(* IEC 61131-3 sources: REFUSR/GP/Refusr.jl/samples (part 4) *)

(* ---- 3-MUX_fives-maven-study.st ---- *)
(*
This code implements a shuffled multiplexer with 3 control bits.
The control bits are: Data[6], Data[2], Data[1]
The input bits are: Data[5], Data[7], Data[8], Data[10], Data[11], Data[9], Data[3], Data[4]

The symbolic expression is:
(((((((~((~(D[6]) & ~(D[2])) & ~(D[1])) | D[5]) & (~((D[6] & ~(D[2])) & ~(D[1])) | D[7])) & (~((~(D[6]) & D[2]) & ~(D[1])) | D[8])) & (~((D[6] & D[2]) & ~(D[1])) | D[10])) & (~((~(D[6]) & ~(D[2])) & D[1]) | D[11])) & (~((D[6] & ~(D[2])) & D[1]) | D[9])) & (~((~(D[6]) & D[2]) & D[1]) | D[3])) & (~((D[6] & D[2]) & D[1]) | D[4])

*)

FUNCTION_BLOCK F_CollectInput
  VAR_IN_OUT
      Data : ARRAY[1..15] OF BOOL;
  END_VAR
  VAR_INPUT
      TICK  : BOOL := 0;
      IN1   : BOOL := 0;
      IN2   : BOOL := 0;
      IN3   : BOOL := 0;
      IN4   : BOOL := 0;
      IN5   : BOOL := 0;
      RESET : BOOL := FALSE;
  END_VAR
  VAR_OUTPUT
      Finished : BOOL;
  END_VAR
  VAR
      j    : USINT := 1;
      tock : BOOL  := 0;
  END_VAR
  IF NOT RESET AND tock = NOT TICK THEN
      Data[j]   := IN1;
      Data[j+1] := IN2;
      Data[j+2] := IN3;
      Data[j+3] := IN4;
      Data[j+4] := IN5;
      j := j + 5;
      tock := TICK;
  ELSE
      j := 1;
      tock := 0;
  END_IF;
  Finished := (j > 15);
END_FUNCTION_BLOCK

PROGRAM Boiler
  VAR
    Data  : ARRAY[1..15] OF BOOL;
    Ready : BOOL;
    CollectInput : F_CollectInput;
  END_VAR
  VAR
    TICK     AT %IX1.0 : BOOL;
    IN1      AT %IX0.3 : BOOL;
    IN2      AT %IX0.4 : BOOL;
    IN3      AT %IX0.5 : BOOL;
    IN4      AT %IX0.6 : BOOL;
    IN5      AT %IX0.7 : BOOL;
    OutReady AT %QX0.0 : BOOL := FALSE;
    FeedNext AT %QX0.1 : BOOL := FALSE;
    Out      AT %QX0.2 : BOOL;
  END_VAR
  CollectInput(TICK:=TICK, IN1:=IN1, IN2:=IN2, IN3:=IN3, IN4:=IN4, IN5:=IN5);
  Ready := CollectInput.Finished;
  FeedNext := 1;
  IF Ready THEN
    Out := (((((((((NOT (((NOT D[6]) AND (NOT D[2])) AND (NOT D[1]))) OR D[5]) AND ((NOT ((D[6] AND (NOT D[2])) AND (NOT D[1]))) OR D[7])) AND ((NOT (((NOT D[6]) AND D[2]) AND (NOT D[1]))) OR D[8])) AND ((NOT ((D[6] AND D[2]) AND (NOT D[1]))) OR D[10])) AND ((NOT (((NOT D[6]) AND (NOT D[2])) AND D[1])) OR D[11])) AND ((NOT ((D[6] AND (NOT D[2])) AND D[1])) OR D[9])) AND ((NOT (((NOT D[6]) AND D[2]) AND D[1])) OR D[3])) AND ((NOT ((D[6] AND D[2]) AND D[1])) OR D[4]));
    OutReady := 1;
    CollectInput(RESET:=TRUE);
  END_IF;
END_PROGRAM

CONFIGURATION Config0
  RESOURCE Res0 ON PLC
    TASK task0(INTERVAL := T#20ms,PRIORITY := 0);
    PROGRAM instance0 WITH task0 : Boiler;
  END_RESOURCE
END_CONFIGURATION

(* ---- 3-MUX_flout-chows-peers.st ---- *)
(*
This code implements a shuffled multiplexer with 3 control bits.
The control bits are: Data[1], Data[2], Data[7]
The input bits are: Data[8], Data[3], Data[5], Data[4], Data[9], Data[6], Data[10], Data[11]

The symbolic expression is:
(((((((~((~(D[1]) & ~(D[2])) & ~(D[7])) | D[8]) & (~((D[1] & ~(D[2])) & ~(D[7])) | D[3])) & (~((~(D[1]) & D[2]) & ~(D[7])) | D[5])) & (~((D[1] & D[2]) & ~(D[7])) | D[4])) & (~((~(D[1]) & ~(D[2])) & D[7]) | D[9])) & (~((D[1] & ~(D[2])) & D[7]) | D[6])) & (~((~(D[1]) & D[2]) & D[7]) | D[10])) & (~((D[1] & D[2]) & D[7]) | D[11])

*)

FUNCTION_BLOCK F_CollectInput
  VAR_IN_OUT
      Data : ARRAY[1..15] OF BOOL;
  END_VAR
  VAR_INPUT
      TICK  : BOOL := 0;
      IN1   : BOOL := 0;
      IN2   : BOOL := 0;
      IN3   : BOOL := 0;
      IN4   : BOOL := 0;
      IN5   : BOOL := 0;
      RESET : BOOL := FALSE;
  END_VAR
  VAR_OUTPUT
      Finished : BOOL;
  END_VAR
  VAR
      j    : USINT := 1;
      tock : BOOL  := 0;
  END_VAR
  IF NOT RESET AND tock = NOT TICK THEN
      Data[j]   := IN1;
      Data[j+1] := IN2;
      Data[j+2] := IN3;
      Data[j+3] := IN4;
      Data[j+4] := IN5;
      j := j + 5;
      tock := TICK;
  ELSE
      j := 1;
      tock := 0;
  END_IF;
  Finished := (j > 15);
END_FUNCTION_BLOCK

PROGRAM Boiler
  VAR
    Data  : ARRAY[1..15] OF BOOL;
    Ready : BOOL;
    CollectInput : F_CollectInput;
  END_VAR
  VAR
    TICK     AT %IX1.0 : BOOL;
    IN1      AT %IX0.3 : BOOL;
    IN2      AT %IX0.4 : BOOL;
    IN3      AT %IX0.5 : BOOL;
    IN4      AT %IX0.6 : BOOL;
    IN5      AT %IX0.7 : BOOL;
    OutReady AT %QX0.0 : BOOL := FALSE;
    FeedNext AT %QX0.1 : BOOL := FALSE;
    Out      AT %QX0.2 : BOOL;
  END_VAR
  CollectInput(TICK:=TICK, IN1:=IN1, IN2:=IN2, IN3:=IN3, IN4:=IN4, IN5:=IN5);
  Ready := CollectInput.Finished;
  FeedNext := 1;
  IF Ready THEN
    Out := (((((((((NOT (((NOT D[1]) AND (NOT D[2])) AND (NOT D[7]))) OR D[8]) AND ((NOT ((D[1] AND (NOT D[2])) AND (NOT D[7]))) OR D[3])) AND ((NOT (((NOT D[1]) AND D[2]) AND (NOT D[7]))) OR D[5])) AND ((NOT ((D[1] AND D[2]) AND (NOT D[7]))) OR D[4])) AND ((NOT (((NOT D[1]) AND (NOT D[2])) AND D[7])) OR D[9])) AND ((NOT ((D[1] AND (NOT D[2])) AND D[7])) OR D[6])) AND ((NOT (((NOT D[1]) AND D[2]) AND D[7])) OR D[10])) AND ((NOT ((D[1] AND D[2]) AND D[7])) OR D[11]));
    OutReady := 1;
    CollectInput(RESET:=TRUE);
  END_IF;
END_PROGRAM

CONFIGURATION Config0
  RESOURCE Res0 ON PLC
    TASK task0(INTERVAL := T#20ms,PRIORITY := 0);
    PROGRAM instance0 WITH task0 : Boiler;
  END_RESOURCE
END_CONFIGURATION

(* ---- 3-MUX_fluff-masse-darts.st ---- *)
(*
This code implements a shuffled multiplexer with 3 control bits.
The control bits are: Data[3], Data[2], Data[1]
The input bits are: Data[5], Data[4], Data[6], Data[9], Data[7], Data[11], Data[10], Data[8]

The symbolic expression is:
(((((((~((~(D[3]) & ~(D[2])) & ~(D[1])) | D[5]) & (~((D[3] & ~(D[2])) & ~(D[1])) | D[4])) & (~((~(D[3]) & D[2]) & ~(D[1])) | D[6])) & (~((D[3] & D[2]) & ~(D[1])) | D[9])) & (~((~(D[3]) & ~(D[2])) & D[1]) | D[7])) & (~((D[3] & ~(D[2])) & D[1]) | D[11])) & (~((~(D[3]) & D[2]) & D[1]) | D[10])) & (~((D[3] & D[2]) & D[1]) | D[8])

*)

FUNCTION_BLOCK F_CollectInput
  VAR_IN_OUT
      Data : ARRAY[1..15] OF BOOL;
  END_VAR
  VAR_INPUT
      TICK  : BOOL := 0;
      IN1   : BOOL := 0;
      IN2   : BOOL := 0;
      IN3   : BOOL := 0;
      IN4   : BOOL := 0;
      IN5   : BOOL := 0;
      RESET : BOOL := FALSE;
  END_VAR
  VAR_OUTPUT
      Finished : BOOL;
  END_VAR
  VAR
      j    : USINT := 1;
      tock : BOOL  := 0;
  END_VAR
  IF NOT RESET AND tock = NOT TICK THEN
      Data[j]   := IN1;
      Data[j+1] := IN2;
      Data[j+2] := IN3;
      Data[j+3] := IN4;
      Data[j+4] := IN5;
      j := j + 5;
      tock := TICK;
  ELSE
      j := 1;
      tock := 0;
  END_IF;
  Finished := (j > 15);
END_FUNCTION_BLOCK

PROGRAM Boiler
  VAR
    Data  : ARRAY[1..15] OF BOOL;
    Ready : BOOL;
    CollectInput : F_CollectInput;
  END_VAR
  VAR
    TICK     AT %IX1.0 : BOOL;
    IN1      AT %IX0.3 : BOOL;
    IN2      AT %IX0.4 : BOOL;
    IN3      AT %IX0.5 : BOOL;
    IN4      AT %IX0.6 : BOOL;
    IN5      AT %IX0.7 : BOOL;
    OutReady AT %QX0.0 : BOOL := FALSE;
    FeedNext AT %QX0.1 : BOOL := FALSE;
    Out      AT %QX0.2 : BOOL;
  END_VAR
  CollectInput(TICK:=TICK, IN1:=IN1, IN2:=IN2, IN3:=IN3, IN4:=IN4, IN5:=IN5);
  Ready := CollectInput.Finished;
  FeedNext := 1;
  IF Ready THEN
    Out := (((((((((NOT (((NOT D[3]) AND (NOT D[2])) AND (NOT D[1]))) OR D[5]) AND ((NOT ((D[3] AND (NOT D[2])) AND (NOT D[1]))) OR D[4])) AND ((NOT (((NOT D[3]) AND D[2]) AND (NOT D[1]))) OR D[6])) AND ((NOT ((D[3] AND D[2]) AND (NOT D[1]))) OR D[9])) AND ((NOT (((NOT D[3]) AND (NOT D[2])) AND D[1])) OR D[7])) AND ((NOT ((D[3] AND (NOT D[2])) AND D[1])) OR D[11])) AND ((NOT (((NOT D[3]) AND D[2]) AND D[1])) OR D[10])) AND ((NOT ((D[3] AND D[2]) AND D[1])) OR D[8]));
    OutReady := 1;
    CollectInput(RESET:=TRUE);
  END_IF;
END_PROGRAM

CONFIGURATION Config0
  RESOURCE Res0 ON PLC
    TASK task0(INTERVAL := T#20ms,PRIORITY := 0);
    PROGRAM instance0 WITH task0 : Boiler;
  END_RESOURCE
END_CONFIGURATION

(* ---- 3-MUX_ftped-surfs-skein.st ---- *)
(*
This code implements a shuffled multiplexer with 3 control bits.
The control bits are: Data[3], Data[2], Data[5]
The input bits are: Data[4], Data[7], Data[8], Data[1], Data[10], Data[6], Data[9], Data[11]

The symbolic expression is:
(((((((~((~(D[3]) & ~(D[2])) & ~(D[5])) | D[4]) & (~((D[3] & ~(D[2])) & ~(D[5])) | D[7])) & (~((~(D[3]) & D[2]) & ~(D[5])) | D[8])) & (~((D[3] & D[2]) & ~(D[5])) | D[1])) & (~((~(D[3]) & ~(D[2])) & D[5]) | D[10])) & (~((D[3] & ~(D[2])) & D[5]) | D[6])) & (~((~(D[3]) & D[2]) & D[5]) | D[9])) & (~((D[3] & D[2]) & D[5]) | D[11])

*)

FUNCTION_BLOCK F_CollectInput
  VAR_IN_OUT
      Data : ARRAY[1..15] OF BOOL;
  END_VAR
  VAR_INPUT
      TICK  : BOOL := 0;
      IN1   : BOOL := 0;
      IN2   : BOOL := 0;
      IN3   : BOOL := 0;
      IN4   : BOOL := 0;
      IN5   : BOOL := 0;
      RESET : BOOL := FALSE;
  END_VAR
  VAR_OUTPUT
      Finished : BOOL;
  END_VAR
  VAR
      j    : USINT := 1;
      tock : BOOL  := 0;
  END_VAR
  IF NOT RESET AND tock = NOT TICK THEN
      Data[j]   := IN1;
      Data[j+1] := IN2;
      Data[j+2] := IN3;
      Data[j+3] := IN4;
      Data[j+4] := IN5;
      j := j + 5;
      tock := TICK;
  ELSE
      j := 1;
      tock := 0;
  END_IF;
  Finished := (j > 15);
END_FUNCTION_BLOCK

PROGRAM Boiler
  VAR
    Data  : ARRAY[1..15] OF BOOL;
    Ready : BOOL;
    CollectInput : F_CollectInput;
  END_VAR
  VAR
    TICK     AT %IX1.0 : BOOL;
    IN1      AT %IX0.3 : BOOL;
    IN2      AT %IX0.4 : BOOL;
    IN3      AT %IX0.5 : BOOL;
    IN4      AT %IX0.6 : BOOL;
    IN5      AT %IX0.7 : BOOL;
    OutReady AT %QX0.0 : BOOL := FALSE;
    FeedNext AT %QX0.1 : BOOL := FALSE;
    Out      AT %QX0.2 : BOOL;
  END_VAR
  CollectInput(TICK:=TICK, IN1:=IN1, IN2:=IN2, IN3:=IN3, IN4:=IN4, IN5:=IN5);
  Ready := CollectInput.Finished;
  FeedNext := 1;
  IF Ready THEN
    Out := (((((((((NOT (((NOT D[3]) AND (NOT D[2])) AND (NOT D[5]))) OR D[4]) AND ((NOT ((D[3] AND (NOT D[2])) AND (NOT D[5]))) OR D[7])) AND ((NOT (((NOT D[3]) AND D[2]) AND (NOT D[5]))) OR D[8])) AND ((NOT ((D[3] AND D[2]) AND (NOT D[5]))) OR D[1])) AND ((NOT (((NOT D[3]) AND (NOT D[2])) AND D[5])) OR D[10])) AND ((NOT ((D[3] AND (NOT D[2])) AND D[5])) OR D[6])) AND ((NOT (((NOT D[3]) AND D[2]) AND D[5])) OR D[9])) AND ((NOT ((D[3] AND D[2]) AND D[5])) OR D[11]));
    OutReady := 1;
    CollectInput(RESET:=TRUE);
  END_IF;
END_PROGRAM

CONFIGURATION Config0
  RESOURCE Res0 ON PLC
    TASK task0(INTERVAL := T#20ms,PRIORITY := 0);
    PROGRAM instance0 WITH task0 : Boiler;
  END_RESOURCE
END_CONFIGURATION

(* ---- 3-MUX_fugal-tawny-pants.st ---- *)
(*
This code implements a shuffled multiplexer with 3 control bits.
The control bits are: Data[1], Data[2], Data[3]
The input bits are: Data[5], Data[9], Data[8], Data[4], Data[10], Data[6], Data[7], Data[11]

The symbolic expression is:
(((((((~((~(D[1]) & ~(D[2])) & ~(D[3])) | D[5]) & (~((D[1] & ~(D[2])) & ~(D[3])) | D[9])) & (~((~(D[1]) & D[2]) & ~(D[3])) | D[8])) & (~((D[1] & D[2]) & ~(D[3])) | D[4])) & (~((~(D[1]) & ~(D[2])) & D[3]) | D[10])) & (~((D[1] & ~(D[2])) & D[3]) | D[6])) & (~((~(D[1]) & D[2]) & D[3]) | D[7])) & (~((D[1] & D[2]) & D[3]) | D[11])

*)

FUNCTION_BLOCK F_CollectInput
  VAR_IN_OUT
      Data : ARRAY[1..15] OF BOOL;
  END_VAR
  VAR_INPUT
      TICK  : BOOL := 0;
      IN1   : BOOL := 0;
      IN2   : BOOL := 0;
      IN3   : BOOL := 0;
      IN4   : BOOL := 0;
      IN5   : BOOL := 0;
      RESET : BOOL := FALSE;
  END_VAR
  VAR_OUTPUT
      Finished : BOOL;
  END_VAR
  VAR
      j    : USINT := 1;
      tock : BOOL  := 0;
  END_VAR
  IF NOT RESET AND tock = NOT TICK THEN
      Data[j]   := IN1;
      Data[j+1] := IN2;
      Data[j+2] := IN3;
      Data[j+3] := IN4;
      Data[j+4] := IN5;
      j := j + 5;
      tock := TICK;
  ELSE
      j := 1;
      tock := 0;
  END_IF;
  Finished := (j > 15);
END_FUNCTION_BLOCK

PROGRAM Boiler
  VAR
    Data  : ARRAY[1..15] OF BOOL;
    Ready : BOOL;
    CollectInput : F_CollectInput;
  END_VAR
  VAR
    TICK     AT %IX1.0 : BOOL;
    IN1      AT %IX0.3 : BOOL;
    IN2      AT %IX0.4 : BOOL;
    IN3      AT %IX0.5 : BOOL;
    IN4      AT %IX0.6 : BOOL;
    IN5      AT %IX0.7 : BOOL;
    OutReady AT %QX0.0 : BOOL := FALSE;
    FeedNext AT %QX0.1 : BOOL := FALSE;
    Out      AT %QX0.2 : BOOL;
  END_VAR
  CollectInput(TICK:=TICK, IN1:=IN1, IN2:=IN2, IN3:=IN3, IN4:=IN4, IN5:=IN5);
  Ready := CollectInput.Finished;
  FeedNext := 1;
  IF Ready THEN
    Out := (((((((((NOT (((NOT D[1]) AND (NOT D[2])) AND (NOT D[3]))) OR D[5]) AND ((NOT ((D[1] AND (NOT D[2])) AND (NOT D[3]))) OR D[9])) AND ((NOT (((NOT D[1]) AND D[2]) AND (NOT D[3]))) OR D[8])) AND ((NOT ((D[1] AND D[2]) AND (NOT D[3]))) OR D[4])) AND ((NOT (((NOT D[1]) AND (NOT D[2])) AND D[3])) OR D[10])) AND ((NOT ((D[1] AND (NOT D[2])) AND D[3])) OR D[6])) AND ((NOT (((NOT D[1]) AND D[2]) AND D[3])) OR D[7])) AND ((NOT ((D[1] AND D[2]) AND D[3])) OR D[11]));
    OutReady := 1;
    CollectInput(RESET:=TRUE);
  END_IF;
END_PROGRAM

CONFIGURATION Config0
  RESOURCE Res0 ON PLC
    TASK task0(INTERVAL := T#20ms,PRIORITY := 0);
    PROGRAM instance0 WITH task0 : Boiler;
  END_RESOURCE
END_CONFIGURATION

(* ---- 3-MUX_ghost-throw-niche.st ---- *)
(*
This code implements a shuffled multiplexer with 3 control bits.
The control bits are: Data[2], Data[1], Data[3]
The input bits are: Data[6], Data[5], Data[7], Data[9], Data[10], Data[4], Data[8], Data[11]

The symbolic expression is:
(((((((~((~(D[2]) & ~(D[1])) & ~(D[3])) | D[6]) & (~((D[2] & ~(D[1])) & ~(D[3])) | D[5])) & (~((~(D[2]) & D[1]) & ~(D[3])) | D[7])) & (~((D[2] & D[1]) & ~(D[3])) | D[9])) & (~((~(D[2]) & ~(D[1])) & D[3]) | D[10])) & (~((D[2] & ~(D[1])) & D[3]) | D[4])) & (~((~(D[2]) & D[1]) & D[3]) | D[8])) & (~((D[2] & D[1]) & D[3]) | D[11])

*)

FUNCTION_BLOCK F_CollectInput
  VAR_IN_OUT
      Data : ARRAY[1..15] OF BOOL;
  END_VAR
  VAR_INPUT
      TICK  : BOOL := 0;
      IN1   : BOOL := 0;
      IN2   : BOOL := 0;
      IN3   : BOOL := 0;
      IN4   : BOOL := 0;
      IN5   : BOOL := 0;
      RESET : BOOL := FALSE;
  END_VAR
  VAR_OUTPUT
      Finished : BOOL;
  END_VAR
  VAR
      j    : USINT := 1;
      tock : BOOL  := 0;
  END_VAR
  IF NOT RESET AND tock = NOT TICK THEN
      Data[j]   := IN1;
      Data[j+1] := IN2;
      Data[j+2] := IN3;
      Data[j+3] := IN4;
      Data[j+4] := IN5;
      j := j + 5;
      tock := TICK;
  ELSE
      j := 1;
      tock := 0;
  END_IF;
  Finished := (j > 15);
END_FUNCTION_BLOCK

PROGRAM Boiler
  VAR
    Data  : ARRAY[1..15] OF BOOL;
    Ready : BOOL;
    CollectInput : F_CollectInput;
  END_VAR
  VAR
    TICK     AT %IX1.0 : BOOL;
    IN1      AT %IX0.3 : BOOL;
    IN2      AT %IX0.4 : BOOL;
    IN3      AT %IX0.5 : BOOL;
    IN4      AT %IX0.6 : BOOL;
    IN5      AT %IX0.7 : BOOL;
    OutReady AT %QX0.0 : BOOL := FALSE;
    FeedNext AT %QX0.1 : BOOL := FALSE;
    Out      AT %QX0.2 : BOOL;
  END_VAR
  CollectInput(TICK:=TICK, IN1:=IN1, IN2:=IN2, IN3:=IN3, IN4:=IN4, IN5:=IN5);
  Ready := CollectInput.Finished;
  FeedNext := 1;
  IF Ready THEN
    Out := (((((((((NOT (((NOT D[2]) AND (NOT D[1])) AND (NOT D[3]))) OR D[6]) AND ((NOT ((D[2] AND (NOT D[1])) AND (NOT D[3]))) OR D[5])) AND ((NOT (((NOT D[2]) AND D[1]) AND (NOT D[3]))) OR D[7])) AND ((NOT ((D[2] AND D[1]) AND (NOT D[3]))) OR D[9])) AND ((NOT (((NOT D[2]) AND (NOT D[1])) AND D[3])) OR D[10])) AND ((NOT ((D[2] AND (NOT D[1])) AND D[3])) OR D[4])) AND ((NOT (((NOT D[2]) AND D[1]) AND D[3])) OR D[8])) AND ((NOT ((D[2] AND D[1]) AND D[3])) OR D[11]));
    OutReady := 1;
    CollectInput(RESET:=TRUE);
  END_IF;
END_PROGRAM

CONFIGURATION Config0
  RESOURCE Res0 ON PLC
    TASK task0(INTERVAL := T#20ms,PRIORITY := 0);
    PROGRAM instance0 WITH task0 : Boiler;
  END_RESOURCE
END_CONFIGURATION

(* ---- 3-MUX_giant-blocs-dicta.st ---- *)
(*
This code implements a shuffled multiplexer with 3 control bits.
The control bits are: Data[1], Data[3], Data[9]
The input bits are: Data[4], Data[2], Data[6], Data[8], Data[7], Data[5], Data[11], Data[10]

The symbolic expression is:
(((((((~((~(D[1]) & ~(D[3])) & ~(D[9])) | D[4]) & (~((D[1] & ~(D[3])) & ~(D[9])) | D[2])) & (~((~(D[1]) & D[3]) & ~(D[9])) | D[6])) & (~((D[1] & D[3]) & ~(D[9])) | D[8])) & (~((~(D[1]) & ~(D[3])) & D[9]) | D[7])) & (~((D[1] & ~(D[3])) & D[9]) | D[5])) & (~((~(D[1]) & D[3]) & D[9]) | D[11])) & (~((D[1] & D[3]) & D[9]) | D[10])

*)

FUNCTION_BLOCK F_CollectInput
  VAR_IN_OUT
      Data : ARRAY[1..15] OF BOOL;
  END_VAR
  VAR_INPUT
      TICK  : BOOL := 0;
      IN1   : BOOL := 0;
      IN2   : BOOL := 0;
      IN3   : BOOL := 0;
      IN4   : BOOL := 0;
      IN5   : BOOL := 0;
      RESET : BOOL := FALSE;
  END_VAR
  VAR_OUTPUT
      Finished : BOOL;
  END_VAR
  VAR
      j    : USINT := 1;
      tock : BOOL  := 0;
  END_VAR
  IF NOT RESET AND tock = NOT TICK THEN
      Data[j]   := IN1;
      Data[j+1] := IN2;
      Data[j+2] := IN3;
      Data[j+3] := IN4;
      Data[j+4] := IN5;
      j := j + 5;
      tock := TICK;
  ELSE
      j := 1;
      tock := 0;
  END_IF;
  Finished := (j > 15);
END_FUNCTION_BLOCK

PROGRAM Boiler
  VAR
    Data  : ARRAY[1..15] OF BOOL;
    Ready : BOOL;
    CollectInput : F_CollectInput;
  END_VAR
  VAR
    TICK     AT %IX1.0 : BOOL;
    IN1      AT %IX0.3 : BOOL;
    IN2      AT %IX0.4 : BOOL;
    IN3      AT %IX0.5 : BOOL;
    IN4      AT %IX0.6 : BOOL;
    IN5      AT %IX0.7 : BOOL;
    OutReady AT %QX0.0 : BOOL := FALSE;
    FeedNext AT %QX0.1 : BOOL := FALSE;
    Out      AT %QX0.2 : BOOL;
  END_VAR
  CollectInput(TICK:=TICK, IN1:=IN1, IN2:=IN2, IN3:=IN3, IN4:=IN4, IN5:=IN5);
  Ready := CollectInput.Finished;
  FeedNext := 1;
  IF Ready THEN
    Out := (((((((((NOT (((NOT D[1]) AND (NOT D[3])) AND (NOT D[9]))) OR D[4]) AND ((NOT ((D[1] AND (NOT D[3])) AND (NOT D[9]))) OR D[2])) AND ((NOT (((NOT D[1]) AND D[3]) AND (NOT D[9]))) OR D[6])) AND ((NOT ((D[1] AND D[3]) AND (NOT D[9]))) OR D[8])) AND ((NOT (((NOT D[1]) AND (NOT D[3])) AND D[9])) OR D[7])) AND ((NOT ((D[1] AND (NOT D[3])) AND D[9])) OR D[5])) AND ((NOT (((NOT D[1]) AND D[3]) AND D[9])) OR D[11])) AND ((NOT ((D[1] AND D[3]) AND D[9])) OR D[10]));
    OutReady := 1;
    CollectInput(RESET:=TRUE);
  END_IF;
END_PROGRAM

CONFIGURATION Config0
  RESOURCE Res0 ON PLC
    TASK task0(INTERVAL := T#20ms,PRIORITY := 0);
    PROGRAM instance0 WITH task0 : Boiler;
  END_RESOURCE
END_CONFIGURATION

(* ---- 3-MUX_goofy-uncap-recap.st ---- *)
(*
This code implements a shuffled multiplexer with 3 control bits.
The control bits are: Data[2], Data[1], Data[4]
The input bits are: Data[3], Data[5], Data[7], Data[6], Data[9], Data[10], Data[11], Data[8]

The symbolic expression is:
(((((((~((~(D[2]) & ~(D[1])) & ~(D[4])) | D[3]) & (~((D[2] & ~(D[1])) & ~(D[4])) | D[5])) & (~((~(D[2]) & D[1]) & ~(D[4])) | D[7])) & (~((D[2] & D[1]) & ~(D[4])) | D[6])) & (~((~(D[2]) & ~(D[1])) & D[4]) | D[9])) & (~((D[2] & ~(D[1])) & D[4]) | D[10])) & (~((~(D[2]) & D[1]) & D[4]) | D[11])) & (~((D[2] & D[1]) & D[4]) | D[8])

*)

FUNCTION_BLOCK F_CollectInput
  VAR_IN_OUT
      Data : ARRAY[1..15] OF BOOL;
  END_VAR
  VAR_INPUT
      TICK  : BOOL := 0;
      IN1   : BOOL := 0;
      IN2   : BOOL := 0;
      IN3   : BOOL := 0;
      IN4   : BOOL := 0;
      IN5   : BOOL := 0;
      RESET : BOOL := FALSE;
  END_VAR
  VAR_OUTPUT
      Finished : BOOL;
  END_VAR
  VAR
      j    : USINT := 1;
      tock : BOOL  := 0;
  END_VAR
  IF NOT RESET AND tock = NOT TICK THEN
      Data[j]   := IN1;
      Data[j+1] := IN2;
      Data[j+2] := IN3;
      Data[j+3] := IN4;
      Data[j+4] := IN5;
      j := j + 5;
      tock := TICK;
  ELSE
      j := 1;
      tock := 0;
  END_IF;
  Finished := (j > 15);
END_FUNCTION_BLOCK

PROGRAM Boiler
  VAR
    Data  : ARRAY[1..15] OF BOOL;
    Ready : BOOL;
    CollectInput : F_CollectInput;
  END_VAR
  VAR
    TICK     AT %IX1.0 : BOOL;
    IN1      AT %IX0.3 : BOOL;
    IN2      AT %IX0.4 : BOOL;
    IN3      AT %IX0.5 : BOOL;
    IN4      AT %IX0.6 : BOOL;
    IN5      AT %IX0.7 : BOOL;
    OutReady AT %QX0.0 : BOOL := FALSE;
    FeedNext AT %QX0.1 : BOOL := FALSE;
    Out      AT %QX0.2 : BOOL;
  END_VAR
  CollectInput(TICK:=TICK, IN1:=IN1, IN2:=IN2, IN3:=IN3, IN4:=IN4, IN5:=IN5);
  Ready := CollectInput.Finished;
  FeedNext := 1;
  IF Ready THEN
    Out := (((((((((NOT (((NOT D[2]) AND (NOT D[1])) AND (NOT D[4]))) OR D[3]) AND ((NOT ((D[2] AND (NOT D[1])) AND (NOT D[4]))) OR D[5])) AND ((NOT (((NOT D[2]) AND D[1]) AND (NOT D[4]))) OR D[7])) AND ((NOT ((D[2] AND D[1]) AND (NOT D[4]))) OR D[6])) AND ((NOT (((NOT D[2]) AND (NOT D[1])) AND D[4])) OR D[9])) AND ((NOT ((D[2] AND (NOT D[1])) AND D[4])) OR D[10])) AND ((NOT (((NOT D[2]) AND D[1]) AND D[4])) OR D[11])) AND ((NOT ((D[2] AND D[1]) AND D[4])) OR D[8]));
    OutReady := 1;
    CollectInput(RESET:=TRUE);
  END_IF;
END_PROGRAM

CONFIGURATION Config0
  RESOURCE Res0 ON PLC
    TASK task0(INTERVAL := T#20ms,PRIORITY := 0);
    PROGRAM instance0 WITH task0 : Boiler;
  END_RESOURCE
END_CONFIGURATION

(* ---- 3-MUX_grunt-trite-rapid.st ---- *)
(*
This code implements a shuffled multiplexer with 3 control bits.
The control bits are: Data[2], Data[3], Data[7]
The input bits are: Data[6], Data[4], Data[1], Data[9], Data[5], Data[10], Data[8], Data[11]

The symbolic expression is:
(((((((~((~(D[2]) & ~(D[3])) & ~(D[7])) | D[6]) & (~((D[2] & ~(D[3])) & ~(D[7])) | D[4])) & (~((~(D[2]) & D[3]) & ~(D[7])) | D[1])) & (~((D[2] & D[3]) & ~(D[7])) | D[9])) & (~((~(D[2]) & ~(D[3])) & D[7]) | D[5])) & (~((D[2] & ~(D[3])) & D[7]) | D[10])) & (~((~(D[2]) & D[3]) & D[7]) | D[8])) & (~((D[2] & D[3]) & D[7]) | D[11])

*)

FUNCTION_BLOCK F_CollectInput
  VAR_IN_OUT
      Data : ARRAY[1..15] OF BOOL;
  END_VAR
  VAR_INPUT
      TICK  : BOOL := 0;
      IN1   : BOOL := 0;
      IN2   : BOOL := 0;
      IN3   : BOOL := 0;
      IN4   : BOOL := 0;
      IN5   : BOOL := 0;
      RESET : BOOL := FALSE;
  END_VAR
  VAR_OUTPUT
      Finished : BOOL;
  END_VAR
  VAR
      j    : USINT := 1;
      tock : BOOL  := 0;
  END_VAR
  IF NOT RESET AND tock = NOT TICK THEN
      Data[j]   := IN1;
      Data[j+1] := IN2;
      Data[j+2] := IN3;
      Data[j+3] := IN4;
      Data[j+4] := IN5;
      j := j + 5;
      tock := TICK;
  ELSE
      j := 1;
      tock := 0;
  END_IF;
  Finished := (j > 15);
END_FUNCTION_BLOCK

PROGRAM Boiler
  VAR
    Data  : ARRAY[1..15] OF BOOL;
    Ready : BOOL;
    CollectInput : F_CollectInput;
  END_VAR
  VAR
    TICK     AT %IX1.0 : BOOL;
    IN1      AT %IX0.3 : BOOL;
    IN2      AT %IX0.4 : BOOL;
    IN3      AT %IX0.5 : BOOL;
    IN4      AT %IX0.6 : BOOL;
    IN5      AT %IX0.7 : BOOL;
    OutReady AT %QX0.0 : BOOL := FALSE;
    FeedNext AT %QX0.1 : BOOL := FALSE;
    Out      AT %QX0.2 : BOOL;
  END_VAR
  CollectInput(TICK:=TICK, IN1:=IN1, IN2:=IN2, IN3:=IN3, IN4:=IN4, IN5:=IN5);
  Ready := CollectInput.Finished;
  FeedNext := 1;
  IF Ready THEN
    Out := (((((((((NOT (((NOT D[2]) AND (NOT D[3])) AND (NOT D[7]))) OR D[6]) AND ((NOT ((D[2] AND (NOT D[3])) AND (NOT D[7]))) OR D[4])) AND ((NOT (((NOT D[2]) AND D[3]) AND (NOT D[7]))) OR D[1])) AND ((NOT ((D[2] AND D[3]) AND (NOT D[7]))) OR D[9])) AND ((NOT (((NOT D[2]) AND (NOT D[3])) AND D[7])) OR D[5])) AND ((NOT ((D[2] AND (NOT D[3])) AND D[7])) OR D[10])) AND ((NOT (((NOT D[2]) AND D[3]) AND D[7])) OR D[8])) AND ((NOT ((D[2] AND D[3]) AND D[7])) OR D[11]));
    OutReady := 1;
    CollectInput(RESET:=TRUE);
  END_IF;
END_PROGRAM

CONFIGURATION Config0
  RESOURCE Res0 ON PLC
    TASK task0(INTERVAL := T#20ms,PRIORITY := 0);
    PROGRAM instance0 WITH task0 : Boiler;
  END_RESOURCE
END_CONFIGURATION

(* ---- 3-MUX_gully-crink-seams.st ---- *)
(*
This code implements a shuffled multiplexer with 3 control bits.
The control bits are: Data[1], Data[3], Data[4]
The input bits are: Data[5], Data[2], Data[6], Data[8], Data[9], Data[10], Data[7], Data[11]

The symbolic expression is:
(((((((~((~(D[1]) & ~(D[3])) & ~(D[4])) | D[5]) & (~((D[1] & ~(D[3])) & ~(D[4])) | D[2])) & (~((~(D[1]) & D[3]) & ~(D[4])) | D[6])) & (~((D[1] & D[3]) & ~(D[4])) | D[8])) & (~((~(D[1]) & ~(D[3])) & D[4]) | D[9])) & (~((D[1] & ~(D[3])) & D[4]) | D[10])) & (~((~(D[1]) & D[3]) & D[4]) | D[7])) & (~((D[1] & D[3]) & D[4]) | D[11])

*)

FUNCTION_BLOCK F_CollectInput
  VAR_IN_OUT
      Data : ARRAY[1..15] OF BOOL;
  END_VAR
  VAR_INPUT
      TICK  : BOOL := 0;
      IN1   : BOOL := 0;
      IN2   : BOOL := 0;
      IN3   : BOOL := 0;
      IN4   : BOOL := 0;
      IN5   : BOOL := 0;
      RESET : BOOL := FALSE;
  END_VAR
  VAR_OUTPUT
      Finished : BOOL;
  END_VAR
  VAR
      j    : USINT := 1;
      tock : BOOL  := 0;
  END_VAR
  IF NOT RESET AND tock = NOT TICK THEN
      Data[j]   := IN1;
      Data[j+1] := IN2;
      Data[j+2] := IN3;
      Data[j+3] := IN4;
      Data[j+4] := IN5;
      j := j + 5;
      tock := TICK;
  ELSE
      j := 1;
      tock := 0;
  END_IF;
  Finished := (j > 15);
END_FUNCTION_BLOCK

PROGRAM Boiler
  VAR
    Data  : ARRAY[1..15] OF BOOL;
    Ready : BOOL;
    CollectInput : F_CollectInput;
  END_VAR
  VAR
    TICK     AT %IX1.0 : BOOL;
    IN1      AT %IX0.3 : BOOL;
    IN2      AT %IX0.4 : BOOL;
    IN3      AT %IX0.5 : BOOL;
    IN4      AT %IX0.6 : BOOL;
    IN5      AT %IX0.7 : BOOL;
    OutReady AT %QX0.0 : BOOL := FALSE;
    FeedNext AT %QX0.1 : BOOL := FALSE;
    Out      AT %QX0.2 : BOOL;
  END_VAR
  CollectInput(TICK:=TICK, IN1:=IN1, IN2:=IN2, IN3:=IN3, IN4:=IN4, IN5:=IN5);
  Ready := CollectInput.Finished;
  FeedNext := 1;
  IF Ready THEN
    Out := (((((((((NOT (((NOT D[1]) AND (NOT D[3])) AND (NOT D[4]))) OR D[5]) AND ((NOT ((D[1] AND (NOT D[3])) AND (NOT D[4]))) OR D[2])) AND ((NOT (((NOT D[1]) AND D[3]) AND (NOT D[4]))) OR D[6])) AND ((NOT ((D[1] AND D[3]) AND (NOT D[4]))) OR D[8])) AND ((NOT (((NOT D[1]) AND (NOT D[3])) AND D[4])) OR D[9])) AND ((NOT ((D[1] AND (NOT D[3])) AND D[4])) OR D[10])) AND ((NOT (((NOT D[1]) AND D[3]) AND D[4])) OR D[7])) AND ((NOT ((D[1] AND D[3]) AND D[4])) OR D[11]));
    OutReady := 1;
    CollectInput(RESET:=TRUE);
  END_IF;
END_PROGRAM

CONFIGURATION Config0
  RESOURCE Res0 ON PLC
    TASK task0(INTERVAL := T#20ms,PRIORITY := 0);
    PROGRAM instance0 WITH task0 : Boiler;
  END_RESOURCE
END_CONFIGURATION

(* ---- 3-MUX_hexes-rumps-hanks.st ---- *)
(*
This code implements a shuffled multiplexer with 3 control bits.
The control bits are: Data[2], Data[3], Data[1]
The input bits are: Data[4], Data[5], Data[8], Data[7], Data[6], Data[9], Data[11], Data[10]

The symbolic expression is:
(((((((~((~(D[2]) & ~(D[3])) & ~(D[1])) | D[4]) & (~((D[2] & ~(D[3])) & ~(D[1])) | D[5])) & (~((~(D[2]) & D[3]) & ~(D[1])) | D[8])) & (~((D[2] & D[3]) & ~(D[1])) | D[7])) & (~((~(D[2]) & ~(D[3])) & D[1]) | D[6])) & (~((D[2] & ~(D[3])) & D[1]) | D[9])) & (~((~(D[2]) & D[3]) & D[1]) | D[11])) & (~((D[2] & D[3]) & D[1]) | D[10])

*)

FUNCTION_BLOCK F_CollectInput
  VAR_IN_OUT
      Data : ARRAY[1..15] OF BOOL;
  END_VAR
  VAR_INPUT
      TICK  : BOOL := 0;
      IN1   : BOOL := 0;
      IN2   : BOOL := 0;
      IN3   : BOOL := 0;
      IN4   : BOOL := 0;
      IN5   : BOOL := 0;
      RESET : BOOL := FALSE;
  END_VAR
  VAR_OUTPUT
      Finished : BOOL;
  END_VAR
  VAR
      j    : USINT := 1;
      tock : BOOL  := 0;
  END_VAR
  IF NOT RESET AND tock = NOT TICK THEN
      Data[j]   := IN1;
      Data[j+1] := IN2;
      Data[j+2] := IN3;
      Data[j+3] := IN4;
      Data[j+4] := IN5;
      j := j + 5;
      tock := TICK;
  ELSE
      j := 1;
      tock := 0;
  END_IF;
  Finished := (j > 15);
END_FUNCTION_BLOCK

PROGRAM Boiler
  VAR
    Data  : ARRAY[1..15] OF BOOL;
    Ready : BOOL;
    CollectInput : F_CollectInput;
  END_VAR
  VAR
    TICK     AT %IX1.0 : BOOL;
    IN1      AT %IX0.3 : BOOL;
    IN2      AT %IX0.4 : BOOL;
    IN3      AT %IX0.5 : BOOL;
    IN4      AT %IX0.6 : BOOL;
    IN5      AT %IX0.7 : BOOL;
    OutReady AT %QX0.0 : BOOL := FALSE;
    FeedNext AT %QX0.1 : BOOL := FALSE;
    Out      AT %QX0.2 : BOOL;
  END_VAR
  CollectInput(TICK:=TICK, IN1:=IN1, IN2:=IN2, IN3:=IN3, IN4:=IN4, IN5:=IN5);
  Ready := CollectInput.Finished;
  FeedNext := 1;
  IF Ready THEN
    Out := (((((((((NOT (((NOT D[2]) AND (NOT D[3])) AND (NOT D[1]))) OR D[4]) AND ((NOT ((D[2] AND (NOT D[3])) AND (NOT D[1]))) OR D[5])) AND ((NOT (((NOT D[2]) AND D[3]) AND (NOT D[1]))) OR D[8])) AND ((NOT ((D[2] AND D[3]) AND (NOT D[1]))) OR D[7])) AND ((NOT (((NOT D[2]) AND (NOT D[3])) AND D[1])) OR D[6])) AND ((NOT ((D[2] AND (NOT D[3])) AND D[1])) OR D[9])) AND ((NOT (((NOT D[2]) AND D[3]) AND D[1])) OR D[11])) AND ((NOT ((D[2] AND D[3]) AND D[1])) OR D[10]));
    OutReady := 1;
    CollectInput(RESET:=TRUE);
  END_IF;
END_PROGRAM

CONFIGURATION Config0
  RESOURCE Res0 ON PLC
    TASK task0(INTERVAL := T#20ms,PRIORITY := 0);
    PROGRAM instance0 WITH task0 : Boiler;
  END_RESOURCE
END_CONFIGURATION

(* ---- 3-MUX_hived-field-nuked.st ---- *)
(*
This code implements a shuffled multiplexer with 3 control bits.
The control bits are: Data[4], Data[3], Data[7]
The input bits are: Data[9], Data[10], Data[1], Data[2], Data[5], Data[6], Data[11], Data[8]

The symbolic expression is:
(((((((~((~(D[4]) & ~(D[3])) & ~(D[7])) | D[9]) & (~((D[4] & ~(D[3])) & ~(D[7])) | D[10])) & (~((~(D[4]) & D[3]) & ~(D[7])) | D[1])) & (~((D[4] & D[3]) & ~(D[7])) | D[2])) & (~((~(D[4]) & ~(D[3])) & D[7]) | D[5])) & (~((D[4] & ~(D[3])) & D[7]) | D[6])) & (~((~(D[4]) & D[3]) & D[7]) | D[11])) & (~((D[4] & D[3]) & D[7]) | D[8])

*)

FUNCTION_BLOCK F_CollectInput
  VAR_IN_OUT
      Data : ARRAY[1..15] OF BOOL;
  END_VAR
  VAR_INPUT
      TICK  : BOOL := 0;
      IN1   : BOOL := 0;
      IN2   : BOOL := 0;
      IN3   : BOOL := 0;
      IN4   : BOOL := 0;
      IN5   : BOOL := 0;
      RESET : BOOL := FALSE;
  END_VAR
  VAR_OUTPUT
      Finished : BOOL;
  END_VAR
  VAR
      j    : USINT := 1;
      tock : BOOL  := 0;
  END_VAR
  IF NOT RESET AND tock = NOT TICK THEN
      Data[j]   := IN1;
      Data[j+1] := IN2;
      Data[j+2] := IN3;
      Data[j+3] := IN4;
      Data[j+4] := IN5;
      j := j + 5;
      tock := TICK;
  ELSE
      j := 1;
      tock := 0;
  END_IF;
  Finished := (j > 15);
END_FUNCTION_BLOCK

PROGRAM Boiler
  VAR
    Data  : ARRAY[1..15] OF BOOL;
    Ready : BOOL;
    CollectInput : F_CollectInput;
  END_VAR
  VAR
    TICK     AT %IX1.0 : BOOL;
    IN1      AT %IX0.3 : BOOL;
    IN2      AT %IX0.4 : BOOL;
    IN3      AT %IX0.5 : BOOL;
    IN4      AT %IX0.6 : BOOL;
    IN5      AT %IX0.7 : BOOL;
    OutReady AT %QX0.0 : BOOL := FALSE;
    FeedNext AT %QX0.1 : BOOL := FALSE;
    Out      AT %QX0.2 : BOOL;
  END_VAR
  CollectInput(TICK:=TICK, IN1:=IN1, IN2:=IN2, IN3:=IN3, IN4:=IN4, IN5:=IN5);
  Ready := CollectInput.Finished;
  FeedNext := 1;
  IF Ready THEN
    Out := (((((((((NOT (((NOT D[4]) AND (NOT D[3])) AND (NOT D[7]))) OR D[9]) AND ((NOT ((D[4] AND (NOT D[3])) AND (NOT D[7]))) OR D[10])) AND ((NOT (((NOT D[4]) AND D[3]) AND (NOT D[7]))) OR D[1])) AND ((NOT ((D[4] AND D[3]) AND (NOT D[7]))) OR D[2])) AND ((NOT (((NOT D[4]) AND (NOT D[3])) AND D[7])) OR D[5])) AND ((NOT ((D[4] AND (NOT D[3])) AND D[7])) OR D[6])) AND ((NOT (((NOT D[4]) AND D[3]) AND D[7])) OR D[11])) AND ((NOT ((D[4] AND D[3]) AND D[7])) OR D[8]));
    OutReady := 1;
    CollectInput(RESET:=TRUE);
  END_IF;
END_PROGRAM

CONFIGURATION Config0
  RESOURCE Res0 ON PLC
    TASK task0(INTERVAL := T#20ms,PRIORITY := 0);
    PROGRAM instance0 WITH task0 : Boiler;
  END_RESOURCE
END_CONFIGURATION

(* ---- 3-MUX_jeeps-bazar-carry.st ---- *)
(*
This code implements a shuffled multiplexer with 3 control bits.
The control bits are: Data[2], Data[1], Data[4]
The input bits are: Data[6], Data[5], Data[3], Data[7], Data[9], Data[8], Data[10], Data[11]

The symbolic expression is:
(((((((~((~(D[2]) & ~(D[1])) & ~(D[4])) | D[6]) & (~((D[2] & ~(D[1])) & ~(D[4])) | D[5])) & (~((~(D[2]) & D[1]) & ~(D[4])) | D[3])) & (~((D[2] & D[1]) & ~(D[4])) | D[7])) & (~((~(D[2]) & ~(D[1])) & D[4]) | D[9])) & (~((D[2] & ~(D[1])) & D[4]) | D[8])) & (~((~(D[2]) & D[1]) & D[4]) | D[10])) & (~((D[2] & D[1]) & D[4]) | D[11])

*)

FUNCTION_BLOCK F_CollectInput
  VAR_IN_OUT
      Data : ARRAY[1..15] OF BOOL;
  END_VAR
  VAR_INPUT
      TICK  : BOOL := 0;
      IN1   : BOOL := 0;
      IN2   : BOOL := 0;
      IN3   : BOOL := 0;
      IN4   : BOOL := 0;
      IN5   : BOOL := 0;
      RESET : BOOL := FALSE;
  END_VAR
  VAR_OUTPUT
      Finished : BOOL;
  END_VAR
  VAR
      j    : USINT := 1;
      tock : BOOL  := 0;
  END_VAR
  IF NOT RESET AND tock = NOT TICK THEN
      Data[j]   := IN1;
      Data[j+1] := IN2;
      Data[j+2] := IN3;
      Data[j+3] := IN4;
      Data[j+4] := IN5;
      j := j + 5;
      tock := TICK;
  ELSE
      j := 1;
      tock := 0;
  END_IF;
  Finished := (j > 15);
END_FUNCTION_BLOCK

PROGRAM Boiler
  VAR
    Data  : ARRAY[1..15] OF BOOL;
    Ready : BOOL;
    CollectInput : F_CollectInput;
  END_VAR
  VAR
    TICK     AT %IX1.0 : BOOL;
    IN1      AT %IX0.3 : BOOL;
    IN2      AT %IX0.4 : BOOL;
    IN3      AT %IX0.5 : BOOL;
    IN4      AT %IX0.6 : BOOL;
    IN5      AT %IX0.7 : BOOL;
    OutReady AT %QX0.0 : BOOL := FALSE;
    FeedNext AT %QX0.1 : BOOL := FALSE;
    Out      AT %QX0.2 : BOOL;
  END_VAR
  CollectInput(TICK:=TICK, IN1:=IN1, IN2:=IN2, IN3:=IN3, IN4:=IN4, IN5:=IN5);
  Ready := CollectInput.Finished;
  FeedNext := 1;
  IF Ready THEN
    Out := (((((((((NOT (((NOT D[2]) AND (NOT D[1])) AND (NOT D[4]))) OR D[6]) AND ((NOT ((D[2] AND (NOT D[1])) AND (NOT D[4]))) OR D[5])) AND ((NOT (((NOT D[2]) AND D[1]) AND (NOT D[4]))) OR D[3])) AND ((NOT ((D[2] AND D[1]) AND (NOT D[4]))) OR D[7])) AND ((NOT (((NOT D[2]) AND (NOT D[1])) AND D[4])) OR D[9])) AND ((NOT ((D[2] AND (NOT D[1])) AND D[4])) OR D[8])) AND ((NOT (((NOT D[2]) AND D[1]) AND D[4])) OR D[10])) AND ((NOT ((D[2] AND D[1]) AND D[4])) OR D[11]));
    OutReady := 1;
    CollectInput(RESET:=TRUE);
  END_IF;
END_PROGRAM

CONFIGURATION Config0
  RESOURCE Res0 ON PLC
    TASK task0(INTERVAL := T#20ms,PRIORITY := 0);
    PROGRAM instance0 WITH task0 : Boiler;
  END_RESOURCE
END_CONFIGURATION

(* ---- 3-MUX_jumps-pussy-stirs.st ---- *)
(*
This code implements a shuffled multiplexer with 3 control bits.
The control bits are: Data[2], Data[3], Data[1]
The input bits are: Data[4], Data[5], Data[8], Data[6], Data[7], Data[9], Data[11], Data[10]

The symbolic expression is:
(((((((~((~(D[2]) & ~(D[3])) & ~(D[1])) | D[4]) & (~((D[2] & ~(D[3])) & ~(D[1])) | D[5])) & (~((~(D[2]) & D[3]) & ~(D[1])) | D[8])) & (~((D[2] & D[3]) & ~(D[1])) | D[6])) & (~((~(D[2]) & ~(D[3])) & D[1]) | D[7])) & (~((D[2] & ~(D[3])) & D[1]) | D[9])) & (~((~(D[2]) & D[3]) & D[1]) | D[11])) & (~((D[2] & D[3]) & D[1]) | D[10])

*)

FUNCTION_BLOCK F_CollectInput
  VAR_IN_OUT
      Data : ARRAY[1..15] OF BOOL;
  END_VAR
  VAR_INPUT
      TICK  : BOOL := 0;
      IN1   : BOOL := 0;
      IN2   : BOOL := 0;
      IN3   : BOOL := 0;
      IN4   : BOOL := 0;
      IN5   : BOOL := 0;
      RESET : BOOL := FALSE;
  END_VAR
  VAR_OUTPUT
      Finished : BOOL;
  END_VAR
  VAR
      j    : USINT := 1;
      tock : BOOL  := 0;
  END_VAR
  IF NOT RESET AND tock = NOT TICK THEN
      Data[j]   := IN1;
      Data[j+1] := IN2;
      Data[j+2] := IN3;
      Data[j+3] := IN4;
      Data[j+4] := IN5;
      j := j + 5;
      tock := TICK;
  ELSE
      j := 1;
      tock := 0;
  END_IF;
  Finished := (j > 15);
END_FUNCTION_BLOCK

PROGRAM Boiler
  VAR
    Data  : ARRAY[1..15] OF BOOL;
    Ready : BOOL;
    CollectInput : F_CollectInput;
  END_VAR
  VAR
    TICK     AT %IX1.0 : BOOL;
    IN1      AT %IX0.3 : BOOL;
    IN2      AT %IX0.4 : BOOL;
    IN3      AT %IX0.5 : BOOL;
    IN4      AT %IX0.6 : BOOL;
    IN5      AT %IX0.7 : BOOL;
    OutReady AT %QX0.0 : BOOL := FALSE;
    FeedNext AT %QX0.1 : BOOL := FALSE;
    Out      AT %QX0.2 : BOOL;
  END_VAR
  CollectInput(TICK:=TICK, IN1:=IN1, IN2:=IN2, IN3:=IN3, IN4:=IN4, IN5:=IN5);
  Ready := CollectInput.Finished;
  FeedNext := 1;
  IF Ready THEN
    Out := (((((((((NOT (((NOT D[2]) AND (NOT D[3])) AND (NOT D[1]))) OR D[4]) AND ((NOT ((D[2] AND (NOT D[3])) AND (NOT D[1]))) OR D[5])) AND ((NOT (((NOT D[2]) AND D[3]) AND (NOT D[1]))) OR D[8])) AND ((NOT ((D[2] AND D[3]) AND (NOT D[1]))) OR D[6])) AND ((NOT (((NOT D[2]) AND (NOT D[3])) AND D[1])) OR D[7])) AND ((NOT ((D[2] AND (NOT D[3])) AND D[1])) OR D[9])) AND ((NOT (((NOT D[2]) AND D[3]) AND D[1])) OR D[11])) AND ((NOT ((D[2] AND D[3]) AND D[1])) OR D[10]));
    OutReady := 1;
    CollectInput(RESET:=TRUE);
  END_IF;
END_PROGRAM

CONFIGURATION Config0
  RESOURCE Res0 ON PLC
    TASK task0(INTERVAL := T#20ms,PRIORITY := 0);
    PROGRAM instance0 WITH task0 : Boiler;
  END_RESOURCE
END_CONFIGURATION

(* ---- 3-MUX_laves-tidal-green.st ---- *)
(*
This code implements a shuffled multiplexer with 3 control bits.
The control bits are: Data[2], Data[3], Data[1]
The input bits are: Data[5], Data[8], Data[6], Data[4], Data[7], Data[9], Data[10], Data[11]

The symbolic expression is:
(((((((~((~(D[2]) & ~(D[3])) & ~(D[1])) | D[5]) & (~((D[2] & ~(D[3])) & ~(D[1])) | D[8])) & (~((~(D[2]) & D[3]) & ~(D[1])) | D[6])) & (~((D[2] & D[3]) & ~(D[1])) | D[4])) & (~((~(D[2]) & ~(D[3])) & D[1]) | D[7])) & (~((D[2] & ~(D[3])) & D[1]) | D[9])) & (~((~(D[2]) & D[3]) & D[1]) | D[10])) & (~((D[2] & D[3]) & D[1]) | D[11])

*)

FUNCTION_BLOCK F_CollectInput
  VAR_IN_OUT
      Data : ARRAY[1..15] OF BOOL;
  END_VAR
  VAR_INPUT
      TICK  : BOOL := 0;
      IN1   : BOOL := 0;
      IN2   : BOOL := 0;
      IN3   : BOOL := 0;
      IN4   : BOOL := 0;
      IN5   : BOOL := 0;
      RESET : BOOL := FALSE;
  END_VAR
  VAR_OUTPUT
      Finished : BOOL;
  END_VAR
  VAR
      j    : USINT := 1;
      tock : BOOL  := 0;
  END_VAR
  IF NOT RESET AND tock = NOT TICK THEN
      Data[j]   := IN1;
      Data[j+1] := IN2;
      Data[j+2] := IN3;
      Data[j+3] := IN4;
      Data[j+4] := IN5;
      j := j + 5;
      tock := TICK;
  ELSE
      j := 1;
      tock := 0;
  END_IF;
  Finished := (j > 15);
END_FUNCTION_BLOCK

PROGRAM Boiler
  VAR
    Data  : ARRAY[1..15] OF BOOL;
    Ready : BOOL;
    CollectInput : F_CollectInput;
  END_VAR
  VAR
    TICK     AT %IX1.0 : BOOL;
    IN1      AT %IX0.3 : BOOL;
    IN2      AT %IX0.4 : BOOL;
    IN3      AT %IX0.5 : BOOL;
    IN4      AT %IX0.6 : BOOL;
    IN5      AT %IX0.7 : BOOL;
    OutReady AT %QX0.0 : BOOL := FALSE;
    FeedNext AT %QX0.1 : BOOL := FALSE;
    Out      AT %QX0.2 : BOOL;
  END_VAR
  CollectInput(TICK:=TICK, IN1:=IN1, IN2:=IN2, IN3:=IN3, IN4:=IN4, IN5:=IN5);
  Ready := CollectInput.Finished;
  FeedNext := 1;
  IF Ready THEN
    Out := (((((((((NOT (((NOT D[2]) AND (NOT D[3])) AND (NOT D[1]))) OR D[5]) AND ((NOT ((D[2] AND (NOT D[3])) AND (NOT D[1]))) OR D[8])) AND ((NOT (((NOT D[2]) AND D[3]) AND (NOT D[1]))) OR D[6])) AND ((NOT ((D[2] AND D[3]) AND (NOT D[1]))) OR D[4])) AND ((NOT (((NOT D[2]) AND (NOT D[3])) AND D[1])) OR D[7])) AND ((NOT ((D[2] AND (NOT D[3])) AND D[1])) OR D[9])) AND ((NOT (((NOT D[2]) AND D[3]) AND D[1])) OR D[10])) AND ((NOT ((D[2] AND D[3]) AND D[1])) OR D[11]));
    OutReady := 1;
    CollectInput(RESET:=TRUE);
  END_IF;
END_PROGRAM

CONFIGURATION Config0
  RESOURCE Res0 ON PLC
    TASK task0(INTERVAL := T#20ms,PRIORITY := 0);
    PROGRAM instance0 WITH task0 : Boiler;
  END_RESOURCE
END_CONFIGURATION

(* ---- 3-MUX_leers-curse-altho.st ---- *)
(*
This code implements a shuffled multiplexer with 3 control bits.
The control bits are: Data[3], Data[1], Data[2]
The input bits are: Data[4], Data[6], Data[5], Data[7], Data[9], Data[8], Data[11], Data[10]

The symbolic expression is:
(((((((~((~(D[3]) & ~(D[1])) & ~(D[2])) | D[4]) & (~((D[3] & ~(D[1])) & ~(D[2])) | D[6])) & (~((~(D[3]) & D[1]) & ~(D[2])) | D[5])) & (~((D[3] & D[1]) & ~(D[2])) | D[7])) & (~((~(D[3]) & ~(D[1])) & D[2]) | D[9])) & (~((D[3] & ~(D[1])) & D[2]) | D[8])) & (~((~(D[3]) & D[1]) & D[2]) | D[11])) & (~((D[3] & D[1]) & D[2]) | D[10])

*)

FUNCTION_BLOCK F_CollectInput
  VAR_IN_OUT
      Data : ARRAY[1..15] OF BOOL;
  END_VAR
  VAR_INPUT
      TICK  : BOOL := 0;
      IN1   : BOOL := 0;
      IN2   : BOOL := 0;
      IN3   : BOOL := 0;
      IN4   : BOOL := 0;
      IN5   : BOOL := 0;
      RESET : BOOL := FALSE;
  END_VAR
  VAR_OUTPUT
      Finished : BOOL;
  END_VAR
  VAR
      j    : USINT := 1;
      tock : BOOL  := 0;
  END_VAR
  IF NOT RESET AND tock = NOT TICK THEN
      Data[j]   := IN1;
      Data[j+1] := IN2;
      Data[j+2] := IN3;
      Data[j+3] := IN4;
      Data[j+4] := IN5;
      j := j + 5;
      tock := TICK;
  ELSE
      j := 1;
      tock := 0;
  END_IF;
  Finished := (j > 15);
END_FUNCTION_BLOCK

PROGRAM Boiler
  VAR
    Data  : ARRAY[1..15] OF BOOL;
    Ready : BOOL;
    CollectInput : F_CollectInput;
  END_VAR
  VAR
    TICK     AT %IX1.0 : BOOL;
    IN1      AT %IX0.3 : BOOL;
    IN2      AT %IX0.4 : BOOL;
    IN3      AT %IX0.5 : BOOL;
    IN4      AT %IX0.6 : BOOL;
    IN5      AT %IX0.7 : BOOL;
    OutReady AT %QX0.0 : BOOL := FALSE;
    FeedNext AT %QX0.1 : BOOL := FALSE;
    Out      AT %QX0.2 : BOOL;
  END_VAR
  CollectInput(TICK:=TICK, IN1:=IN1, IN2:=IN2, IN3:=IN3, IN4:=IN4, IN5:=IN5);
  Ready := CollectInput.Finished;
  FeedNext := 1;
  IF Ready THEN
    Out := (((((((((NOT (((NOT D[3]) AND (NOT D[1])) AND (NOT D[2]))) OR D[4]) AND ((NOT ((D[3] AND (NOT D[1])) AND (NOT D[2]))) OR D[6])) AND ((NOT (((NOT D[3]) AND D[1]) AND (NOT D[2]))) OR D[5])) AND ((NOT ((D[3] AND D[1]) AND (NOT D[2]))) OR D[7])) AND ((NOT (((NOT D[3]) AND (NOT D[1])) AND D[2])) OR D[9])) AND ((NOT ((D[3] AND (NOT D[1])) AND D[2])) OR D[8])) AND ((NOT (((NOT D[3]) AND D[1]) AND D[2])) OR D[11])) AND ((NOT ((D[3] AND D[1]) AND D[2])) OR D[10]));
    OutReady := 1;
    CollectInput(RESET:=TRUE);
  END_IF;
END_PROGRAM

CONFIGURATION Config0
  RESOURCE Res0 ON PLC
    TASK task0(INTERVAL := T#20ms,PRIORITY := 0);
    PROGRAM instance0 WITH task0 : Boiler;
  END_RESOURCE
END_CONFIGURATION

(* ---- 3-MUX_legos-taker-gauze.st ---- *)
(*
This code implements a shuffled multiplexer with 3 control bits.
The control bits are: Data[2], Data[1], Data[3]
The input bits are: Data[6], Data[5], Data[7], Data[4], Data[8], Data[9], Data[11], Data[10]

The symbolic expression is:
(((((((~((~(D[2]) & ~(D[1])) & ~(D[3])) | D[6]) & (~((D[2] & ~(D[1])) & ~(D[3])) | D[5])) & (~((~(D[2]) & D[1]) & ~(D[3])) | D[7])) & (~((D[2] & D[1]) & ~(D[3])) | D[4])) & (~((~(D[2]) & ~(D[1])) & D[3]) | D[8])) & (~((D[2] & ~(D[1])) & D[3]) | D[9])) & (~((~(D[2]) & D[1]) & D[3]) | D[11])) & (~((D[2] & D[1]) & D[3]) | D[10])

*)

FUNCTION_BLOCK F_CollectInput
  VAR_IN_OUT
      Data : ARRAY[1..15] OF BOOL;
  END_VAR
  VAR_INPUT
      TICK  : BOOL := 0;
      IN1   : BOOL := 0;
      IN2   : BOOL := 0;
      IN3   : BOOL := 0;
      IN4   : BOOL := 0;
      IN5   : BOOL := 0;
      RESET : BOOL := FALSE;
  END_VAR
  VAR_OUTPUT
      Finished : BOOL;
  END_VAR
  VAR
      j    : USINT := 1;
      tock : BOOL  := 0;
  END_VAR
  IF NOT RESET AND tock = NOT TICK THEN
      Data[j]   := IN1;
      Data[j+1] := IN2;
      Data[j+2] := IN3;
      Data[j+3] := IN4;
      Data[j+4] := IN5;
      j := j + 5;
      tock := TICK;
  ELSE
      j := 1;
      tock := 0;
  END_IF;
  Finished := (j > 15);
END_FUNCTION_BLOCK

PROGRAM Boiler
  VAR
    Data  : ARRAY[1..15] OF BOOL;
    Ready : BOOL;
    CollectInput : F_CollectInput;
  END_VAR
  VAR
    TICK     AT %IX1.0 : BOOL;
    IN1      AT %IX0.3 : BOOL;
    IN2      AT %IX0.4 : BOOL;
    IN3      AT %IX0.5 : BOOL;
    IN4      AT %IX0.6 : BOOL;
    IN5      AT %IX0.7 : BOOL;
    OutReady AT %QX0.0 : BOOL := FALSE;
    FeedNext AT %QX0.1 : BOOL := FALSE;
    Out      AT %QX0.2 : BOOL;
  END_VAR
  CollectInput(TICK:=TICK, IN1:=IN1, IN2:=IN2, IN3:=IN3, IN4:=IN4, IN5:=IN5);
  Ready := CollectInput.Finished;
  FeedNext := 1;
  IF Ready THEN
    Out := (((((((((NOT (((NOT D[2]) AND (NOT D[1])) AND (NOT D[3]))) OR D[6]) AND ((NOT ((D[2] AND (NOT D[1])) AND (NOT D[3]))) OR D[5])) AND ((NOT (((NOT D[2]) AND D[1]) AND (NOT D[3]))) OR D[7])) AND ((NOT ((D[2] AND D[1]) AND (NOT D[3]))) OR D[4])) AND ((NOT (((NOT D[2]) AND (NOT D[1])) AND D[3])) OR D[8])) AND ((NOT ((D[2] AND (NOT D[1])) AND D[3])) OR D[9])) AND ((NOT (((NOT D[2]) AND D[1]) AND D[3])) OR D[11])) AND ((NOT ((D[2] AND D[1]) AND D[3])) OR D[10]));
    OutReady := 1;
    CollectInput(RESET:=TRUE);
  END_IF;
END_PROGRAM

CONFIGURATION Config0
  RESOURCE Res0 ON PLC
    TASK task0(INTERVAL := T#20ms,PRIORITY := 0);
    PROGRAM instance0 WITH task0 : Boiler;
  END_RESOURCE
END_CONFIGURATION

(* ---- 3-MUX_loony-spume-duvet.st ---- *)
(*
This code implements a shuffled multiplexer with 3 control bits.
The control bits are: Data[1], Data[2], Data[3]
The input bits are: Data[5], Data[6], Data[10], Data[4], Data[11], Data[7], Data[8], Data[9]

The symbolic expression is:
(((((((~((~(D[1]) & ~(D[2])) & ~(D[3])) | D[5]) & (~((D[1] & ~(D[2])) & ~(D[3])) | D[6])) & (~((~(D[1]) & D[2]) & ~(D[3])) | D[10])) & (~((D[1] & D[2]) & ~(D[3])) | D[4])) & (~((~(D[1]) & ~(D[2])) & D[3]) | D[11])) & (~((D[1] & ~(D[2])) & D[3]) | D[7])) & (~((~(D[1]) & D[2]) & D[3]) | D[8])) & (~((D[1] & D[2]) & D[3]) | D[9])

*)

FUNCTION_BLOCK F_CollectInput
  VAR_IN_OUT
      Data : ARRAY[1..15] OF BOOL;
  END_VAR
  VAR_INPUT
      TICK  : BOOL := 0;
      IN1   : BOOL := 0;
      IN2   : BOOL := 0;
      IN3   : BOOL := 0;
      IN4   : BOOL := 0;
      IN5   : BOOL := 0;
      RESET : BOOL := FALSE;
  END_VAR
  VAR_OUTPUT
      Finished : BOOL;
  END_VAR
  VAR
      j    : USINT := 1;
      tock : BOOL  := 0;
  END_VAR
  IF NOT RESET AND tock = NOT TICK THEN
      Data[j]   := IN1;
      Data[j+1] := IN2;
      Data[j+2] := IN3;
      Data[j+3] := IN4;
      Data[j+4] := IN5;
      j := j + 5;
      tock := TICK;
  ELSE
      j := 1;
      tock := 0;
  END_IF;
  Finished := (j > 15);
END_FUNCTION_BLOCK

PROGRAM Boiler
  VAR
    Data  : ARRAY[1..15] OF BOOL;
    Ready : BOOL;
    CollectInput : F_CollectInput;
  END_VAR
  VAR
    TICK     AT %IX1.0 : BOOL;
    IN1      AT %IX0.3 : BOOL;
    IN2      AT %IX0.4 : BOOL;
    IN3      AT %IX0.5 : BOOL;
    IN4      AT %IX0.6 : BOOL;
    IN5      AT %IX0.7 : BOOL;
    OutReady AT %QX0.0 : BOOL := FALSE;
    FeedNext AT %QX0.1 : BOOL := FALSE;
    Out      AT %QX0.2 : BOOL;
  END_VAR
  CollectInput(TICK:=TICK, IN1:=IN1, IN2:=IN2, IN3:=IN3, IN4:=IN4, IN5:=IN5);
  Ready := CollectInput.Finished;
  FeedNext := 1;
  IF Ready THEN
    Out := (((((((((NOT (((NOT D[1]) AND (NOT D[2])) AND (NOT D[3]))) OR D[5]) AND ((NOT ((D[1] AND (NOT D[2])) AND (NOT D[3]))) OR D[6])) AND ((NOT (((NOT D[1]) AND D[2]) AND (NOT D[3]))) OR D[10])) AND ((NOT ((D[1] AND D[2]) AND (NOT D[3]))) OR D[4])) AND ((NOT (((NOT D[1]) AND (NOT D[2])) AND D[3])) OR D[11])) AND ((NOT ((D[1] AND (NOT D[2])) AND D[3])) OR D[7])) AND ((NOT (((NOT D[1]) AND D[2]) AND D[3])) OR D[8])) AND ((NOT ((D[1] AND D[2]) AND D[3])) OR D[9]));
    OutReady := 1;
    CollectInput(RESET:=TRUE);
  END_IF;
END_PROGRAM

CONFIGURATION Config0
  RESOURCE Res0 ON PLC
    TASK task0(INTERVAL := T#20ms,PRIORITY := 0);
    PROGRAM instance0 WITH task0 : Boiler;
  END_RESOURCE
END_CONFIGURATION

(* ---- 3-MUX_magus-taxol-cones.st ---- *)
(*
This code implements a shuffled multiplexer with 3 control bits.
The control bits are: Data[3], Data[2], Data[4]
The input bits are: Data[1], Data[6], Data[5], Data[8], Data[7], Data[9], Data[10], Data[11]

The symbolic expression is:
(((((((~((~(D[3]) & ~(D[2])) & ~(D[4])) | D[1]) & (~((D[3] & ~(D[2])) & ~(D[4])) | D[6])) & (~((~(D[3]) & D[2]) & ~(D[4])) | D[5])) & (~((D[3] & D[2]) & ~(D[4])) | D[8])) & (~((~(D[3]) & ~(D[2])) & D[4]) | D[7])) & (~((D[3] & ~(D[2])) & D[4]) | D[9])) & (~((~(D[3]) & D[2]) & D[4]) | D[10])) & (~((D[3] & D[2]) & D[4]) | D[11])

*)

FUNCTION_BLOCK F_CollectInput
  VAR_IN_OUT
      Data : ARRAY[1..15] OF BOOL;
  END_VAR
  VAR_INPUT
      TICK  : BOOL := 0;
      IN1   : BOOL := 0;
      IN2   : BOOL := 0;
      IN3   : BOOL := 0;
      IN4   : BOOL := 0;
      IN5   : BOOL := 0;
      RESET : BOOL := FALSE;
  END_VAR
  VAR_OUTPUT
      Finished : BOOL;
  END_VAR
  VAR
      j    : USINT := 1;
      tock : BOOL  := 0;
  END_VAR
  IF NOT RESET AND tock = NOT TICK THEN
      Data[j]   := IN1;
      Data[j+1] := IN2;
      Data[j+2] := IN3;
      Data[j+3] := IN4;
      Data[j+4] := IN5;
      j := j + 5;
      tock := TICK;
  ELSE
      j := 1;
      tock := 0;
  END_IF;
  Finished := (j > 15);
END_FUNCTION_BLOCK

PROGRAM Boiler
  VAR
    Data  : ARRAY[1..15] OF BOOL;
    Ready : BOOL;
    CollectInput : F_CollectInput;
  END_VAR
  VAR
    TICK     AT %IX1.0 : BOOL;
    IN1      AT %IX0.3 : BOOL;
    IN2      AT %IX0.4 : BOOL;
    IN3      AT %IX0.5 : BOOL;
    IN4      AT %IX0.6 : BOOL;
    IN5      AT %IX0.7 : BOOL;
    OutReady AT %QX0.0 : BOOL := FALSE;
    FeedNext AT %QX0.1 : BOOL := FALSE;
    Out      AT %QX0.2 : BOOL;
  END_VAR
  CollectInput(TICK:=TICK, IN1:=IN1, IN2:=IN2, IN3:=IN3, IN4:=IN4, IN5:=IN5);
  Ready := CollectInput.Finished;
  FeedNext := 1;
  IF Ready THEN
    Out := (((((((((NOT (((NOT D[3]) AND (NOT D[2])) AND (NOT D[4]))) OR D[1]) AND ((NOT ((D[3] AND (NOT D[2])) AND (NOT D[4]))) OR D[6])) AND ((NOT (((NOT D[3]) AND D[2]) AND (NOT D[4]))) OR D[5])) AND ((NOT ((D[3] AND D[2]) AND (NOT D[4]))) OR D[8])) AND ((NOT (((NOT D[3]) AND (NOT D[2])) AND D[4])) OR D[7])) AND ((NOT ((D[3] AND (NOT D[2])) AND D[4])) OR D[9])) AND ((NOT (((NOT D[3]) AND D[2]) AND D[4])) OR D[10])) AND ((NOT ((D[3] AND D[2]) AND D[4])) OR D[11]));
    OutReady := 1;
    CollectInput(RESET:=TRUE);
  END_IF;
END_PROGRAM

CONFIGURATION Config0
  RESOURCE Res0 ON PLC
    TASK task0(INTERVAL := T#20ms,PRIORITY := 0);
    PROGRAM instance0 WITH task0 : Boiler;
  END_RESOURCE
END_CONFIGURATION

(* ---- 3-MUX_mazes-villi-eared.st ---- *)
(*
This code implements a shuffled multiplexer with 3 control bits.
The control bits are: Data[8], Data[3], Data[4]
The input bits are: Data[2], Data[1], Data[5], Data[6], Data[7], Data[9], Data[10], Data[11]

The symbolic expression is:
(((((((~((~(D[8]) & ~(D[3])) & ~(D[4])) | D[2]) & (~((D[8] & ~(D[3])) & ~(D[4])) | D[1])) & (~((~(D[8]) & D[3]) & ~(D[4])) | D[5])) & (~((D[8] & D[3]) & ~(D[4])) | D[6])) & (~((~(D[8]) & ~(D[3])) & D[4]) | D[7])) & (~((D[8] & ~(D[3])) & D[4]) | D[9])) & (~((~(D[8]) & D[3]) & D[4]) | D[10])) & (~((D[8] & D[3]) & D[4]) | D[11])

*)

FUNCTION_BLOCK F_CollectInput
  VAR_IN_OUT
      Data : ARRAY[1..15] OF BOOL;
  END_VAR
  VAR_INPUT
      TICK  : BOOL := 0;
      IN1   : BOOL := 0;
      IN2   : BOOL := 0;
      IN3   : BOOL := 0;
      IN4   : BOOL := 0;
      IN5   : BOOL := 0;
      RESET : BOOL := FALSE;
  END_VAR
  VAR_OUTPUT
      Finished : BOOL;
  END_VAR
  VAR
      j    : USINT := 1;
      tock : BOOL  := 0;
  END_VAR
  IF NOT RESET AND tock = NOT TICK THEN
      Data[j]   := IN1;
      Data[j+1] := IN2;
      Data[j+2] := IN3;
      Data[j+3] := IN4;
      Data[j+4] := IN5;
      j := j + 5;
      tock := TICK;
  ELSE
      j := 1;
      tock := 0;
  END_IF;
  Finished := (j > 15);
END_FUNCTION_BLOCK

PROGRAM Boiler
  VAR
    Data  : ARRAY[1..15] OF BOOL;
    Ready : BOOL;
    CollectInput : F_CollectInput;
  END_VAR
  VAR
    TICK     AT %IX1.0 : BOOL;
    IN1      AT %IX0.3 : BOOL;
    IN2      AT %IX0.4 : BOOL;
    IN3      AT %IX0.5 : BOOL;
    IN4      AT %IX0.6 : BOOL;
    IN5      AT %IX0.7 : BOOL;
    OutReady AT %QX0.0 : BOOL := FALSE;
    FeedNext AT %QX0.1 : BOOL := FALSE;
    Out      AT %QX0.2 : BOOL;
  END_VAR
  CollectInput(TICK:=TICK, IN1:=IN1, IN2:=IN2, IN3:=IN3, IN4:=IN4, IN5:=IN5);
  Ready := CollectInput.Finished;
  FeedNext := 1;
  IF Ready THEN
    Out := (((((((((NOT (((NOT D[8]) AND (NOT D[3])) AND (NOT D[4]))) OR D[2]) AND ((NOT ((D[8] AND (NOT D[3])) AND (NOT D[4]))) OR D[1])) AND ((NOT (((NOT D[8]) AND D[3]) AND (NOT D[4]))) OR D[5])) AND ((NOT ((D[8] AND D[3]) AND (NOT D[4]))) OR D[6])) AND ((NOT (((NOT D[8]) AND (NOT D[3])) AND D[4])) OR D[7])) AND ((NOT ((D[8] AND (NOT D[3])) AND D[4])) OR D[9])) AND ((NOT (((NOT D[8]) AND D[3]) AND D[4])) OR D[10])) AND ((NOT ((D[8] AND D[3]) AND D[4])) OR D[11]));
    OutReady := 1;
    CollectInput(RESET:=TRUE);
  END_IF;
END_PROGRAM

CONFIGURATION Config0
  RESOURCE Res0 ON PLC
    TASK task0(INTERVAL := T#20ms,PRIORITY := 0);
    PROGRAM instance0 WITH task0 : Boiler;
  END_RESOURCE
END_CONFIGURATION

(* ---- 3-MUX_meaty-inane-flush.st ---- *)
(*
This code implements a shuffled multiplexer with 3 control bits.
The control bits are: Data[2], Data[1], Data[4]
The input bits are: Data[3], Data[6], Data[9], Data[11], Data[7], Data[5], Data[8], Data[10]

The symbolic expression is:
(((((((~((~(D[2]) & ~(D[1])) & ~(D[4])) | D[3]) & (~((D[2] & ~(D[1])) & ~(D[4])) | D[6])) & (~((~(D[2]) & D[1]) & ~(D[4])) | D[9])) & (~((D[2] & D[1]) & ~(D[4])) | D[11])) & (~((~(D[2]) & ~(D[1])) & D[4]) | D[7])) & (~((D[2] & ~(D[1])) & D[4]) | D[5])) & (~((~(D[2]) & D[1]) & D[4]) | D[8])) & (~((D[2] & D[1]) & D[4]) | D[10])

*)

FUNCTION_BLOCK F_CollectInput
  VAR_IN_OUT
      Data : ARRAY[1..15] OF BOOL;
  END_VAR
  VAR_INPUT
      TICK  : BOOL := 0;
      IN1   : BOOL := 0;
      IN2   : BOOL := 0;
      IN3   : BOOL := 0;
      IN4   : BOOL := 0;
      IN5   : BOOL := 0;
      RESET : BOOL := FALSE;
  END_VAR
  VAR_OUTPUT
      Finished : BOOL;
  END_VAR
  VAR
      j    : USINT := 1;
      tock : BOOL  := 0;
  END_VAR
  IF NOT RESET AND tock = NOT TICK THEN
      Data[j]   := IN1;
      Data[j+1] := IN2;
      Data[j+2] := IN3;
      Data[j+3] := IN4;
      Data[j+4] := IN5;
      j := j + 5;
      tock := TICK;
  ELSE
      j := 1;
      tock := 0;
  END_IF;
  Finished := (j > 15);
END_FUNCTION_BLOCK

PROGRAM Boiler
  VAR
    Data  : ARRAY[1..15] OF BOOL;
    Ready : BOOL;
    CollectInput : F_CollectInput;
  END_VAR
  VAR
    TICK     AT %IX1.0 : BOOL;
    IN1      AT %IX0.3 : BOOL;
    IN2      AT %IX0.4 : BOOL;
    IN3      AT %IX0.5 : BOOL;
    IN4      AT %IX0.6 : BOOL;
    IN5      AT %IX0.7 : BOOL;
    OutReady AT %QX0.0 : BOOL := FALSE;
    FeedNext AT %QX0.1 : BOOL := FALSE;
    Out      AT %QX0.2 : BOOL;
  END_VAR
  CollectInput(TICK:=TICK, IN1:=IN1, IN2:=IN2, IN3:=IN3, IN4:=IN4, IN5:=IN5);
  Ready := CollectInput.Finished;
  FeedNext := 1;
  IF Ready THEN
    Out := (((((((((NOT (((NOT D[2]) AND (NOT D[1])) AND (NOT D[4]))) OR D[3]) AND ((NOT ((D[2] AND (NOT D[1])) AND (NOT D[4]))) OR D[6])) AND ((NOT (((NOT D[2]) AND D[1]) AND (NOT D[4]))) OR D[9])) AND ((NOT ((D[2] AND D[1]) AND (NOT D[4]))) OR D[11])) AND ((NOT (((NOT D[2]) AND (NOT D[1])) AND D[4])) OR D[7])) AND ((NOT ((D[2] AND (NOT D[1])) AND D[4])) OR D[5])) AND ((NOT (((NOT D[2]) AND D[1]) AND D[4])) OR D[8])) AND ((NOT ((D[2] AND D[1]) AND D[4])) OR D[10]));
    OutReady := 1;
    CollectInput(RESET:=TRUE);
  END_IF;
END_PROGRAM

CONFIGURATION Config0
  RESOURCE Res0 ON PLC
    TASK task0(INTERVAL := T#20ms,PRIORITY := 0);
    PROGRAM instance0 WITH task0 : Boiler;
  END_RESOURCE
END_CONFIGURATION

(* ---- 3-MUX_melba-snuff-cried.st ---- *)
(*
This code implements a shuffled multiplexer with 3 control bits.
The control bits are: Data[3], Data[1], Data[4]
The input bits are: Data[9], Data[5], Data[10], Data[2], Data[6], Data[7], Data[11], Data[8]

The symbolic expression is:
(((((((~((~(D[3]) & ~(D[1])) & ~(D[4])) | D[9]) & (~((D[3] & ~(D[1])) & ~(D[4])) | D[5])) & (~((~(D[3]) & D[1]) & ~(D[4])) | D[10])) & (~((D[3] & D[1]) & ~(D[4])) | D[2])) & (~((~(D[3]) & ~(D[1])) & D[4]) | D[6])) & (~((D[3] & ~(D[1])) & D[4]) | D[7])) & (~((~(D[3]) & D[1]) & D[4]) | D[11])) & (~((D[3] & D[1]) & D[4]) | D[8])

*)

FUNCTION_BLOCK F_CollectInput
  VAR_IN_OUT
      Data : ARRAY[1..15] OF BOOL;
  END_VAR
  VAR_INPUT
      TICK  : BOOL := 0;
      IN1   : BOOL := 0;
      IN2   : BOOL := 0;
      IN3   : BOOL := 0;
      IN4   : BOOL := 0;
      IN5   : BOOL := 0;
      RESET : BOOL := FALSE;
  END_VAR
  VAR_OUTPUT
      Finished : BOOL;
  END_VAR
  VAR
      j    : USINT := 1;
      tock : BOOL  := 0;
  END_VAR
  IF NOT RESET AND tock = NOT TICK THEN
      Data[j]   := IN1;
      Data[j+1] := IN2;
      Data[j+2] := IN3;
      Data[j+3] := IN4;
      Data[j+4] := IN5;
      j := j + 5;
      tock := TICK;
  ELSE
      j := 1;
      tock := 0;
  END_IF;
  Finished := (j > 15);
END_FUNCTION_BLOCK

PROGRAM Boiler
  VAR
    Data  : ARRAY[1..15] OF BOOL;
    Ready : BOOL;
    CollectInput : F_CollectInput;
  END_VAR
  VAR
    TICK     AT %IX1.0 : BOOL;
    IN1      AT %IX0.3 : BOOL;
    IN2      AT %IX0.4 : BOOL;
    IN3      AT %IX0.5 : BOOL;
    IN4      AT %IX0.6 : BOOL;
    IN5      AT %IX0.7 : BOOL;
    OutReady AT %QX0.0 : BOOL := FALSE;
    FeedNext AT %QX0.1 : BOOL := FALSE;
    Out      AT %QX0.2 : BOOL;
  END_VAR
  CollectInput(TICK:=TICK, IN1:=IN1, IN2:=IN2, IN3:=IN3, IN4:=IN4, IN5:=IN5);
  Ready := CollectInput.Finished;
  FeedNext := 1;
  IF Ready THEN
    Out := (((((((((NOT (((NOT D[3]) AND (NOT D[1])) AND (NOT D[4]))) OR D[9]) AND ((NOT ((D[3] AND (NOT D[1])) AND (NOT D[4]))) OR D[5])) AND ((NOT (((NOT D[3]) AND D[1]) AND (NOT D[4]))) OR D[10])) AND ((NOT ((D[3] AND D[1]) AND (NOT D[4]))) OR D[2])) AND ((NOT (((NOT D[3]) AND (NOT D[1])) AND D[4])) OR D[6])) AND ((NOT ((D[3] AND (NOT D[1])) AND D[4])) OR D[7])) AND ((NOT (((NOT D[3]) AND D[1]) AND D[4])) OR D[11])) AND ((NOT ((D[3] AND D[1]) AND D[4])) OR D[8]));
    OutReady := 1;
    CollectInput(RESET:=TRUE);
  END_IF;
END_PROGRAM

CONFIGURATION Config0
  RESOURCE Res0 ON PLC
    TASK task0(INTERVAL := T#20ms,PRIORITY := 0);
    PROGRAM instance0 WITH task0 : Boiler;
  END_RESOURCE
END_CONFIGURATION

(* ---- 3-MUX_miens-lance-mazer.st ---- *)
(*
This code implements a shuffled multiplexer with 3 control bits.
The control bits are: Data[3], Data[2], Data[1]
The input bits are: Data[4], Data[5], Data[7], Data[6], Data[8], Data[10], Data[9], Data[11]

The symbolic expression is:
(((((((~((~(D[3]) & ~(D[2])) & ~(D[1])) | D[4]) & (~((D[3] & ~(D[2])) & ~(D[1])) | D[5])) & (~((~(D[3]) & D[2]) & ~(D[1])) | D[7])) & (~((D[3] & D[2]) & ~(D[1])) | D[6])) & (~((~(D[3]) & ~(D[2])) & D[1]) | D[8])) & (~((D[3] & ~(D[2])) & D[1]) | D[10])) & (~((~(D[3]) & D[2]) & D[1]) | D[9])) & (~((D[3] & D[2]) & D[1]) | D[11])

*)

FUNCTION_BLOCK F_CollectInput
  VAR_IN_OUT
      Data : ARRAY[1..15] OF BOOL;
  END_VAR
  VAR_INPUT
      TICK  : BOOL := 0;
      IN1   : BOOL := 0;
      IN2   : BOOL := 0;
      IN3   : BOOL := 0;
      IN4   : BOOL := 0;
      IN5   : BOOL := 0;
      RESET : BOOL := FALSE;
  END_VAR
  VAR_OUTPUT
      Finished : BOOL;
  END_VAR
  VAR
      j    : USINT := 1;
      tock : BOOL  := 0;
  END_VAR
  IF NOT RESET AND tock = NOT TICK THEN
      Data[j]   := IN1;
      Data[j+1] := IN2;
      Data[j+2] := IN3;
      Data[j+3] := IN4;
      Data[j+4] := IN5;
      j := j + 5;
      tock := TICK;
  ELSE
      j := 1;
      tock := 0;
  END_IF;
  Finished := (j > 15);
END_FUNCTION_BLOCK

PROGRAM Boiler
  VAR
    Data  : ARRAY[1..15] OF BOOL;
    Ready : BOOL;
    CollectInput : F_CollectInput;
  END_VAR
  VAR
    TICK     AT %IX1.0 : BOOL;
    IN1      AT %IX0.3 : BOOL;
    IN2      AT %IX0.4 : BOOL;
    IN3      AT %IX0.5 : BOOL;
    IN4      AT %IX0.6 : BOOL;
    IN5      AT %IX0.7 : BOOL;
    OutReady AT %QX0.0 : BOOL := FALSE;
    FeedNext AT %QX0.1 : BOOL := FALSE;
    Out      AT %QX0.2 : BOOL;
  END_VAR
  CollectInput(TICK:=TICK, IN1:=IN1, IN2:=IN2, IN3:=IN3, IN4:=IN4, IN5:=IN5);
  Ready := CollectInput.Finished;
  FeedNext := 1;
  IF Ready THEN
    Out := (((((((((NOT (((NOT D[3]) AND (NOT D[2])) AND (NOT D[1]))) OR D[4]) AND ((NOT ((D[3] AND (NOT D[2])) AND (NOT D[1]))) OR D[5])) AND ((NOT (((NOT D[3]) AND D[2]) AND (NOT D[1]))) OR D[7])) AND ((NOT ((D[3] AND D[2]) AND (NOT D[1]))) OR D[6])) AND ((NOT (((NOT D[3]) AND (NOT D[2])) AND D[1])) OR D[8])) AND ((NOT ((D[3] AND (NOT D[2])) AND D[1])) OR D[10])) AND ((NOT (((NOT D[3]) AND D[2]) AND D[1])) OR D[9])) AND ((NOT ((D[3] AND D[2]) AND D[1])) OR D[11]));
    OutReady := 1;
    CollectInput(RESET:=TRUE);
  END_IF;
END_PROGRAM

CONFIGURATION Config0
  RESOURCE Res0 ON PLC
    TASK task0(INTERVAL := T#20ms,PRIORITY := 0);
    PROGRAM instance0 WITH task0 : Boiler;
  END_RESOURCE
END_CONFIGURATION

(* ---- 3-MUX_mints-wicks-ruled.st ---- *)
(*
This code implements a shuffled multiplexer with 3 control bits.
The control bits are: Data[4], Data[2], Data[1]
The input bits are: Data[3], Data[5], Data[7], Data[10], Data[6], Data[9], Data[8], Data[11]

The symbolic expression is:
(((((((~((~(D[4]) & ~(D[2])) & ~(D[1])) | D[3]) & (~((D[4] & ~(D[2])) & ~(D[1])) | D[5])) & (~((~(D[4]) & D[2]) & ~(D[1])) | D[7])) & (~((D[4] & D[2]) & ~(D[1])) | D[10])) & (~((~(D[4]) & ~(D[2])) & D[1]) | D[6])) & (~((D[4] & ~(D[2])) & D[1]) | D[9])) & (~((~(D[4]) & D[2]) & D[1]) | D[8])) & (~((D[4] & D[2]) & D[1]) | D[11])

*)

FUNCTION_BLOCK F_CollectInput
  VAR_IN_OUT
      Data : ARRAY[1..15] OF BOOL;
  END_VAR
  VAR_INPUT
      TICK  : BOOL := 0;
      IN1   : BOOL := 0;
      IN2   : BOOL := 0;
      IN3   : BOOL := 0;
      IN4   : BOOL := 0;
      IN5   : BOOL := 0;
      RESET : BOOL := FALSE;
  END_VAR
  VAR_OUTPUT
      Finished : BOOL;
  END_VAR
  VAR
      j    : USINT := 1;
      tock : BOOL  := 0;
  END_VAR
  IF NOT RESET AND tock = NOT TICK THEN
      Data[j]   := IN1;
      Data[j+1] := IN2;
      Data[j+2] := IN3;
      Data[j+3] := IN4;
      Data[j+4] := IN5;
      j := j + 5;
      tock := TICK;
  ELSE
      j := 1;
      tock := 0;
  END_IF;
  Finished := (j > 15);
END_FUNCTION_BLOCK

PROGRAM Boiler
  VAR
    Data  : ARRAY[1..15] OF BOOL;
    Ready : BOOL;
    CollectInput : F_CollectInput;
  END_VAR
  VAR
    TICK     AT %IX1.0 : BOOL;
    IN1      AT %IX0.3 : BOOL;
    IN2      AT %IX0.4 : BOOL;
    IN3      AT %IX0.5 : BOOL;
    IN4      AT %IX0.6 : BOOL;
    IN5      AT %IX0.7 : BOOL;
    OutReady AT %QX0.0 : BOOL := FALSE;
    FeedNext AT %QX0.1 : BOOL := FALSE;
    Out      AT %QX0.2 : BOOL;
  END_VAR
  CollectInput(TICK:=TICK, IN1:=IN1, IN2:=IN2, IN3:=IN3, IN4:=IN4, IN5:=IN5);
  Ready := CollectInput.Finished;
  FeedNext := 1;
  IF Ready THEN
    Out := (((((((((NOT (((NOT D[4]) AND (NOT D[2])) AND (NOT D[1]))) OR D[3]) AND ((NOT ((D[4] AND (NOT D[2])) AND (NOT D[1]))) OR D[5])) AND ((NOT (((NOT D[4]) AND D[2]) AND (NOT D[1]))) OR D[7])) AND ((NOT ((D[4] AND D[2]) AND (NOT D[1]))) OR D[10])) AND ((NOT (((NOT D[4]) AND (NOT D[2])) AND D[1])) OR D[6])) AND ((NOT ((D[4] AND (NOT D[2])) AND D[1])) OR D[9])) AND ((NOT (((NOT D[4]) AND D[2]) AND D[1])) OR D[8])) AND ((NOT ((D[4] AND D[2]) AND D[1])) OR D[11]));
    OutReady := 1;
    CollectInput(RESET:=TRUE);
  END_IF;
END_PROGRAM

CONFIGURATION Config0
  RESOURCE Res0 ON PLC
    TASK task0(INTERVAL := T#20ms,PRIORITY := 0);
    PROGRAM instance0 WITH task0 : Boiler;
  END_RESOURCE
END_CONFIGURATION

(* ---- 3-MUX_molar-beret-quint.st ---- *)
(*
This code implements a shuffled multiplexer with 3 control bits.
The control bits are: Data[1], Data[2], Data[3]
The input bits are: Data[7], Data[4], Data[5], Data[6], Data[9], Data[8], Data[10], Data[11]

The symbolic expression is:
(((((((~((~(D[1]) & ~(D[2])) & ~(D[3])) | D[7]) & (~((D[1] & ~(D[2])) & ~(D[3])) | D[4])) & (~((~(D[1]) & D[2]) & ~(D[3])) | D[5])) & (~((D[1] & D[2]) & ~(D[3])) | D[6])) & (~((~(D[1]) & ~(D[2])) & D[3]) | D[9])) & (~((D[1] & ~(D[2])) & D[3]) | D[8])) & (~((~(D[1]) & D[2]) & D[3]) | D[10])) & (~((D[1] & D[2]) & D[3]) | D[11])

*)

FUNCTION_BLOCK F_CollectInput
  VAR_IN_OUT
      Data : ARRAY[1..15] OF BOOL;
  END_VAR
  VAR_INPUT
      TICK  : BOOL := 0;
      IN1   : BOOL := 0;
      IN2   : BOOL := 0;
      IN3   : BOOL := 0;
      IN4   : BOOL := 0;
      IN5   : BOOL := 0;
      RESET : BOOL := FALSE;
  END_VAR
  VAR_OUTPUT
      Finished : BOOL;
  END_VAR
  VAR
      j    : USINT := 1;
      tock : BOOL  := 0;
  END_VAR
  IF NOT RESET AND tock = NOT TICK THEN
      Data[j]   := IN1;
      Data[j+1] := IN2;
      Data[j+2] := IN3;
      Data[j+3] := IN4;
      Data[j+4] := IN5;
      j := j + 5;
      tock := TICK;
  ELSE
      j := 1;
      tock := 0;
  END_IF;
  Finished := (j > 15);
END_FUNCTION_BLOCK

PROGRAM Boiler
  VAR
    Data  : ARRAY[1..15] OF BOOL;
    Ready : BOOL;
    CollectInput : F_CollectInput;
  END_VAR
  VAR
    TICK     AT %IX1.0 : BOOL;
    IN1      AT %IX0.3 : BOOL;
    IN2      AT %IX0.4 : BOOL;
    IN3      AT %IX0.5 : BOOL;
    IN4      AT %IX0.6 : BOOL;
    IN5      AT %IX0.7 : BOOL;
    OutReady AT %QX0.0 : BOOL := FALSE;
    FeedNext AT %QX0.1 : BOOL := FALSE;
    Out      AT %QX0.2 : BOOL;
  END_VAR
  CollectInput(TICK:=TICK, IN1:=IN1, IN2:=IN2, IN3:=IN3, IN4:=IN4, IN5:=IN5);
  Ready := CollectInput.Finished;
  FeedNext := 1;
  IF Ready THEN
    Out := (((((((((NOT (((NOT D[1]) AND (NOT D[2])) AND (NOT D[3]))) OR D[7]) AND ((NOT ((D[1] AND (NOT D[2])) AND (NOT D[3]))) OR D[4])) AND ((NOT (((NOT D[1]) AND D[2]) AND (NOT D[3]))) OR D[5])) AND ((NOT ((D[1] AND D[2]) AND (NOT D[3]))) OR D[6])) AND ((NOT (((NOT D[1]) AND (NOT D[2])) AND D[3])) OR D[9])) AND ((NOT ((D[1] AND (NOT D[2])) AND D[3])) OR D[8])) AND ((NOT (((NOT D[1]) AND D[2]) AND D[3])) OR D[10])) AND ((NOT ((D[1] AND D[2]) AND D[3])) OR D[11]));
    OutReady := 1;
    CollectInput(RESET:=TRUE);
  END_IF;
END_PROGRAM

CONFIGURATION Config0
  RESOURCE Res0 ON PLC
    TASK task0(INTERVAL := T#20ms,PRIORITY := 0);
    PROGRAM instance0 WITH task0 : Boiler;
  END_RESOURCE
END_CONFIGURATION

(* ---- 3-MUX_noise-pulps-drubs.st ---- *)
(*
This code implements a shuffled multiplexer with 3 control bits.
The control bits are: Data[1], Data[2], Data[3]
The input bits are: Data[7], Data[6], Data[4], Data[10], Data[8], Data[5], Data[9], Data[11]

The symbolic expression is:
(((((((~((~(D[1]) & ~(D[2])) & ~(D[3])) | D[7]) & (~((D[1] & ~(D[2])) & ~(D[3])) | D[6])) & (~((~(D[1]) & D[2]) & ~(D[3])) | D[4])) & (~((D[1] & D[2]) & ~(D[3])) | D[10])) & (~((~(D[1]) & ~(D[2])) & D[3]) | D[8])) & (~((D[1] & ~(D[2])) & D[3]) | D[5])) & (~((~(D[1]) & D[2]) & D[3]) | D[9])) & (~((D[1] & D[2]) & D[3]) | D[11])

*)

FUNCTION_BLOCK F_CollectInput
  VAR_IN_OUT
      Data : ARRAY[1..15] OF BOOL;
  END_VAR
  VAR_INPUT
      TICK  : BOOL := 0;
      IN1   : BOOL := 0;
      IN2   : BOOL := 0;
      IN3   : BOOL := 0;
      IN4   : BOOL := 0;
      IN5   : BOOL := 0;
      RESET : BOOL := FALSE;
  END_VAR
  VAR_OUTPUT
      Finished : BOOL;
  END_VAR
  VAR
      j    : USINT := 1;
      tock : BOOL  := 0;
  END_VAR
  IF NOT RESET AND tock = NOT TICK THEN
      Data[j]   := IN1;
      Data[j+1] := IN2;
      Data[j+2] := IN3;
      Data[j+3] := IN4;
      Data[j+4] := IN5;
      j := j + 5;
      tock := TICK;
  ELSE
      j := 1;
      tock := 0;
  END_IF;
  Finished := (j > 15);
END_FUNCTION_BLOCK

PROGRAM Boiler
  VAR
    Data  : ARRAY[1..15] OF BOOL;
    Ready : BOOL;
    CollectInput : F_CollectInput;
  END_VAR
  VAR
    TICK     AT %IX1.0 : BOOL;
    IN1      AT %IX0.3 : BOOL;
    IN2      AT %IX0.4 : BOOL;
    IN3      AT %IX0.5 : BOOL;
    IN4      AT %IX0.6 : BOOL;
    IN5      AT %IX0.7 : BOOL;
    OutReady AT %QX0.0 : BOOL := FALSE;
    FeedNext AT %QX0.1 : BOOL := FALSE;
    Out      AT %QX0.2 : BOOL;
  END_VAR
  CollectInput(TICK:=TICK, IN1:=IN1, IN2:=IN2, IN3:=IN3, IN4:=IN4, IN5:=IN5);
  Ready := CollectInput.Finished;
  FeedNext := 1;
  IF Ready THEN
    Out := (((((((((NOT (((NOT D[1]) AND (NOT D[2])) AND (NOT D[3]))) OR D[7]) AND ((NOT ((D[1] AND (NOT D[2])) AND (NOT D[3]))) OR D[6])) AND ((NOT (((NOT D[1]) AND D[2]) AND (NOT D[3]))) OR D[4])) AND ((NOT ((D[1] AND D[2]) AND (NOT D[3]))) OR D[10])) AND ((NOT (((NOT D[1]) AND (NOT D[2])) AND D[3])) OR D[8])) AND ((NOT ((D[1] AND (NOT D[2])) AND D[3])) OR D[5])) AND ((NOT (((NOT D[1]) AND D[2]) AND D[3])) OR D[9])) AND ((NOT ((D[1] AND D[2]) AND D[3])) OR D[11]));
    OutReady := 1;
    CollectInput(RESET:=TRUE);
  END_IF;
END_PROGRAM

CONFIGURATION Config0
  RESOURCE Res0 ON PLC
    TASK task0(INTERVAL := T#20ms,PRIORITY := 0);
    PROGRAM instance0 WITH task0 : Boiler;
  END_RESOURCE
END_CONFIGURATION

(* ---- 3-MUX_omens-fuses-geese.st ---- *)
(*
This code implements a shuffled multiplexer with 3 control bits.
The control bits are: Data[1], Data[3], Data[4]
The input bits are: Data[2], Data[5], Data[6], Data[9], Data[8], Data[7], Data[10], Data[11]

The symbolic expression is:
(((((((~((~(D[1]) & ~(D[3])) & ~(D[4])) | D[2]) & (~((D[1] & ~(D[3])) & ~(D[4])) | D[5])) & (~((~(D[1]) & D[3]) & ~(D[4])) | D[6])) & (~((D[1] & D[3]) & ~(D[4])) | D[9])) & (~((~(D[1]) & ~(D[3])) & D[4]) | D[8])) & (~((D[1] & ~(D[3])) & D[4]) | D[7])) & (~((~(D[1]) & D[3]) & D[4]) | D[10])) & (~((D[1] & D[3]) & D[4]) | D[11])

*)

FUNCTION_BLOCK F_CollectInput
  VAR_IN_OUT
      Data : ARRAY[1..15] OF BOOL;
  END_VAR
  VAR_INPUT
      TICK  : BOOL := 0;
      IN1   : BOOL := 0;
      IN2   : BOOL := 0;
      IN3   : BOOL := 0;
      IN4   : BOOL := 0;
      IN5   : BOOL := 0;
      RESET : BOOL := FALSE;
  END_VAR
  VAR_OUTPUT
      Finished : BOOL;
  END_VAR
  VAR
      j    : USINT := 1;
      tock : BOOL  := 0;
  END_VAR
  IF NOT RESET AND tock = NOT TICK THEN
      Data[j]   := IN1;
      Data[j+1] := IN2;
      Data[j+2] := IN3;
      Data[j+3] := IN4;
      Data[j+4] := IN5;
      j := j + 5;
      tock := TICK;
  ELSE
      j := 1;
      tock := 0;
  END_IF;
  Finished := (j > 15);
END_FUNCTION_BLOCK

PROGRAM Boiler
  VAR
    Data  : ARRAY[1..15] OF BOOL;
    Ready : BOOL;
    CollectInput : F_CollectInput;
  END_VAR
  VAR
    TICK     AT %IX1.0 : BOOL;
    IN1      AT %IX0.3 : BOOL;
    IN2      AT %IX0.4 : BOOL;
    IN3      AT %IX0.5 : BOOL;
    IN4      AT %IX0.6 : BOOL;
    IN5      AT %IX0.7 : BOOL;
    OutReady AT %QX0.0 : BOOL := FALSE;
    FeedNext AT %QX0.1 : BOOL := FALSE;
    Out      AT %QX0.2 : BOOL;
  END_VAR
  CollectInput(TICK:=TICK, IN1:=IN1, IN2:=IN2, IN3:=IN3, IN4:=IN4, IN5:=IN5);
  Ready := CollectInput.Finished;
  FeedNext := 1;
  IF Ready THEN
    Out := (((((((((NOT (((NOT D[1]) AND (NOT D[3])) AND (NOT D[4]))) OR D[2]) AND ((NOT ((D[1] AND (NOT D[3])) AND (NOT D[4]))) OR D[5])) AND ((NOT (((NOT D[1]) AND D[3]) AND (NOT D[4]))) OR D[6])) AND ((NOT ((D[1] AND D[3]) AND (NOT D[4]))) OR D[9])) AND ((NOT (((NOT D[1]) AND (NOT D[3])) AND D[4])) OR D[8])) AND ((NOT ((D[1] AND (NOT D[3])) AND D[4])) OR D[7])) AND ((NOT (((NOT D[1]) AND D[3]) AND D[4])) OR D[10])) AND ((NOT ((D[1] AND D[3]) AND D[4])) OR D[11]));
    OutReady := 1;
    CollectInput(RESET:=TRUE);
  END_IF;
END_PROGRAM

CONFIGURATION Config0
  RESOURCE Res0 ON PLC
    TASK task0(INTERVAL := T#20ms,PRIORITY := 0);
    PROGRAM instance0 WITH task0 : Boiler;
  END_RESOURCE
END_CONFIGURATION

(* ---- 3-MUX_paren-wrier-early.st ---- *)
(*
This code implements a shuffled multiplexer with 3 control bits.
The control bits are: Data[3], Data[1], Data[2]
The input bits are: Data[5], Data[9], Data[4], Data[6], Data[7], Data[8], Data[11], Data[10]

The symbolic expression is:
(((((((~((~(D[3]) & ~(D[1])) & ~(D[2])) | D[5]) & (~((D[3] & ~(D[1])) & ~(D[2])) | D[9])) & (~((~(D[3]) & D[1]) & ~(D[2])) | D[4])) & (~((D[3] & D[1]) & ~(D[2])) | D[6])) & (~((~(D[3]) & ~(D[1])) & D[2]) | D[7])) & (~((D[3] & ~(D[1])) & D[2]) | D[8])) & (~((~(D[3]) & D[1]) & D[2]) | D[11])) & (~((D[3] & D[1]) & D[2]) | D[10])

*)

FUNCTION_BLOCK F_CollectInput
  VAR_IN_OUT
      Data : ARRAY[1..15] OF BOOL;
  END_VAR
  VAR_INPUT
      TICK  : BOOL := 0;
      IN1   : BOOL := 0;
      IN2   : BOOL := 0;
      IN3   : BOOL := 0;
      IN4   : BOOL := 0;
      IN5   : BOOL := 0;
      RESET : BOOL := FALSE;
  END_VAR
  VAR_OUTPUT
      Finished : BOOL;
  END_VAR
  VAR
      j    : USINT := 1;
      tock : BOOL  := 0;
  END_VAR
  IF NOT RESET AND tock = NOT TICK THEN
      Data[j]   := IN1;
      Data[j+1] := IN2;
      Data[j+2] := IN3;
      Data[j+3] := IN4;
      Data[j+4] := IN5;
      j := j + 5;
      tock := TICK;
  ELSE
      j := 1;
      tock := 0;
  END_IF;
  Finished := (j > 15);
END_FUNCTION_BLOCK

PROGRAM Boiler
  VAR
    Data  : ARRAY[1..15] OF BOOL;
    Ready : BOOL;
    CollectInput : F_CollectInput;
  END_VAR
  VAR
    TICK     AT %IX1.0 : BOOL;
    IN1      AT %IX0.3 : BOOL;
    IN2      AT %IX0.4 : BOOL;
    IN3      AT %IX0.5 : BOOL;
    IN4      AT %IX0.6 : BOOL;
    IN5      AT %IX0.7 : BOOL;
    OutReady AT %QX0.0 : BOOL := FALSE;
    FeedNext AT %QX0.1 : BOOL := FALSE;
    Out      AT %QX0.2 : BOOL;
  END_VAR
  CollectInput(TICK:=TICK, IN1:=IN1, IN2:=IN2, IN3:=IN3, IN4:=IN4, IN5:=IN5);
  Ready := CollectInput.Finished;
  FeedNext := 1;
  IF Ready THEN
    Out := (((((((((NOT (((NOT D[3]) AND (NOT D[1])) AND (NOT D[2]))) OR D[5]) AND ((NOT ((D[3] AND (NOT D[1])) AND (NOT D[2]))) OR D[9])) AND ((NOT (((NOT D[3]) AND D[1]) AND (NOT D[2]))) OR D[4])) AND ((NOT ((D[3] AND D[1]) AND (NOT D[2]))) OR D[6])) AND ((NOT (((NOT D[3]) AND (NOT D[1])) AND D[2])) OR D[7])) AND ((NOT ((D[3] AND (NOT D[1])) AND D[2])) OR D[8])) AND ((NOT (((NOT D[3]) AND D[1]) AND D[2])) OR D[11])) AND ((NOT ((D[3] AND D[1]) AND D[2])) OR D[10]));
    OutReady := 1;
    CollectInput(RESET:=TRUE);
  END_IF;
END_PROGRAM

CONFIGURATION Config0
  RESOURCE Res0 ON PLC
    TASK task0(INTERVAL := T#20ms,PRIORITY := 0);
    PROGRAM instance0 WITH task0 : Boiler;
  END_RESOURCE
END_CONFIGURATION

(* ---- 3-MUX_parts-locus-thyme.st ---- *)
(*
This code implements a shuffled multiplexer with 3 control bits.
The control bits are: Data[2], Data[1], Data[5]
The input bits are: Data[3], Data[4], Data[7], Data[6], Data[8], Data[10], Data[9], Data[11]

The symbolic expression is:
(((((((~((~(D[2]) & ~(D[1])) & ~(D[5])) | D[3]) & (~((D[2] & ~(D[1])) & ~(D[5])) | D[4])) & (~((~(D[2]) & D[1]) & ~(D[5])) | D[7])) & (~((D[2] & D[1]) & ~(D[5])) | D[6])) & (~((~(D[2]) & ~(D[1])) & D[5]) | D[8])) & (~((D[2] & ~(D[1])) & D[5]) | D[10])) & (~((~(D[2]) & D[1]) & D[5]) | D[9])) & (~((D[2] & D[1]) & D[5]) | D[11])

*)

FUNCTION_BLOCK F_CollectInput
  VAR_IN_OUT
      Data : ARRAY[1..15] OF BOOL;
  END_VAR
  VAR_INPUT
      TICK  : BOOL := 0;
      IN1   : BOOL := 0;
      IN2   : BOOL := 0;
      IN3   : BOOL := 0;
      IN4   : BOOL := 0;
      IN5   : BOOL := 0;
      RESET : BOOL := FALSE;
  END_VAR
  VAR_OUTPUT
      Finished : BOOL;
  END_VAR
  VAR
      j    : USINT := 1;
      tock : BOOL  := 0;
  END_VAR
  IF NOT RESET AND tock = NOT TICK THEN
      Data[j]   := IN1;
      Data[j+1] := IN2;
      Data[j+2] := IN3;
      Data[j+3] := IN4;
      Data[j+4] := IN5;
      j := j + 5;
      tock := TICK;
  ELSE
      j := 1;
      tock := 0;
  END_IF;
  Finished := (j > 15);
END_FUNCTION_BLOCK

PROGRAM Boiler
  VAR
    Data  : ARRAY[1..15] OF BOOL;
    Ready : BOOL;
    CollectInput : F_CollectInput;
  END_VAR
  VAR
    TICK     AT %IX1.0 : BOOL;
    IN1      AT %IX0.3 : BOOL;
    IN2      AT %IX0.4 : BOOL;
    IN3      AT %IX0.5 : BOOL;
    IN4      AT %IX0.6 : BOOL;
    IN5      AT %IX0.7 : BOOL;
    OutReady AT %QX0.0 : BOOL := FALSE;
    FeedNext AT %QX0.1 : BOOL := FALSE;
    Out      AT %QX0.2 : BOOL;
  END_VAR
  CollectInput(TICK:=TICK, IN1:=IN1, IN2:=IN2, IN3:=IN3, IN4:=IN4, IN5:=IN5);
  Ready := CollectInput.Finished;
  FeedNext := 1;
  IF Ready THEN
    Out := (((((((((NOT (((NOT D[2]) AND (NOT D[1])) AND (NOT D[5]))) OR D[3]) AND ((NOT ((D[2] AND (NOT D[1])) AND (NOT D[5]))) OR D[4])) AND ((NOT (((NOT D[2]) AND D[1]) AND (NOT D[5]))) OR D[7])) AND ((NOT ((D[2] AND D[1]) AND (NOT D[5]))) OR D[6])) AND ((NOT (((NOT D[2]) AND (NOT D[1])) AND D[5])) OR D[8])) AND ((NOT ((D[2] AND (NOT D[1])) AND D[5])) OR D[10])) AND ((NOT (((NOT D[2]) AND D[1]) AND D[5])) OR D[9])) AND ((NOT ((D[2] AND D[1]) AND D[5])) OR D[11]));
    OutReady := 1;
    CollectInput(RESET:=TRUE);
  END_IF;
END_PROGRAM

CONFIGURATION Config0
  RESOURCE Res0 ON PLC
    TASK task0(INTERVAL := T#20ms,PRIORITY := 0);
    PROGRAM instance0 WITH task0 : Boiler;
  END_RESOURCE
END_CONFIGURATION

(* ---- 3-MUX_peals-never-lance.st ---- *)
(*
This code implements a shuffled multiplexer with 3 control bits.
The control bits are: Data[3], Data[2], Data[1]
The input bits are: Data[4], Data[5], Data[6], Data[7], Data[10], Data[8], Data[9], Data[11]

The symbolic expression is:
(((((((~((~(D[3]) & ~(D[2])) & ~(D[1])) | D[4]) & (~((D[3] & ~(D[2])) & ~(D[1])) | D[5])) & (~((~(D[3]) & D[2]) & ~(D[1])) | D[6])) & (~((D[3] & D[2]) & ~(D[1])) | D[7])) & (~((~(D[3]) & ~(D[2])) & D[1]) | D[10])) & (~((D[3] & ~(D[2])) & D[1]) | D[8])) & (~((~(D[3]) & D[2]) & D[1]) | D[9])) & (~((D[3] & D[2]) & D[1]) | D[11])

*)

FUNCTION_BLOCK F_CollectInput
  VAR_IN_OUT
      Data : ARRAY[1..15] OF BOOL;
  END_VAR
  VAR_INPUT
      TICK  : BOOL := 0;
      IN1   : BOOL := 0;
      IN2   : BOOL := 0;
      IN3   : BOOL := 0;
      IN4   : BOOL := 0;
      IN5   : BOOL := 0;
      RESET : BOOL := FALSE;
  END_VAR
  VAR_OUTPUT
      Finished : BOOL;
  END_VAR
  VAR
      j    : USINT := 1;
      tock : BOOL  := 0;
  END_VAR
  IF NOT RESET AND tock = NOT TICK THEN
      Data[j]   := IN1;
      Data[j+1] := IN2;
      Data[j+2] := IN3;
      Data[j+3] := IN4;
      Data[j+4] := IN5;
      j := j + 5;
      tock := TICK;
  ELSE
      j := 1;
      tock := 0;
  END_IF;
  Finished := (j > 15);
END_FUNCTION_BLOCK

PROGRAM Boiler
  VAR
    Data  : ARRAY[1..15] OF BOOL;
    Ready : BOOL;
    CollectInput : F_CollectInput;
  END_VAR
  VAR
    TICK     AT %IX1.0 : BOOL;
    IN1      AT %IX0.3 : BOOL;
    IN2      AT %IX0.4 : BOOL;
    IN3      AT %IX0.5 : BOOL;
    IN4      AT %IX0.6 : BOOL;
    IN5      AT %IX0.7 : BOOL;
    OutReady AT %QX0.0 : BOOL := FALSE;
    FeedNext AT %QX0.1 : BOOL := FALSE;
    Out      AT %QX0.2 : BOOL;
  END_VAR
  CollectInput(TICK:=TICK, IN1:=IN1, IN2:=IN2, IN3:=IN3, IN4:=IN4, IN5:=IN5);
  Ready := CollectInput.Finished;
  FeedNext := 1;
  IF Ready THEN
    Out := (((((((((NOT (((NOT D[3]) AND (NOT D[2])) AND (NOT D[1]))) OR D[4]) AND ((NOT ((D[3] AND (NOT D[2])) AND (NOT D[1]))) OR D[5])) AND ((NOT (((NOT D[3]) AND D[2]) AND (NOT D[1]))) OR D[6])) AND ((NOT ((D[3] AND D[2]) AND (NOT D[1]))) OR D[7])) AND ((NOT (((NOT D[3]) AND (NOT D[2])) AND D[1])) OR D[10])) AND ((NOT ((D[3] AND (NOT D[2])) AND D[1])) OR D[8])) AND ((NOT (((NOT D[3]) AND D[2]) AND D[1])) OR D[9])) AND ((NOT ((D[3] AND D[2]) AND D[1])) OR D[11]));
    OutReady := 1;
    CollectInput(RESET:=TRUE);
  END_IF;
END_PROGRAM

CONFIGURATION Config0
  RESOURCE Res0 ON PLC
    TASK task0(INTERVAL := T#20ms,PRIORITY := 0);
    PROGRAM instance0 WITH task0 : Boiler;
  END_RESOURCE
END_CONFIGURATION

(* ---- 3-MUX_phage-moose-lepta.st ---- *)
(*
This code implements a shuffled multiplexer with 3 control bits.
The control bits are: Data[3], Data[1], Data[4]
The input bits are: Data[5], Data[2], Data[7], Data[8], Data[6], Data[10], Data[11], Data[9]

The symbolic expression is:
(((((((~((~(D[3]) & ~(D[1])) & ~(D[4])) | D[5]) & (~((D[3] & ~(D[1])) & ~(D[4])) | D[2])) & (~((~(D[3]) & D[1]) & ~(D[4])) | D[7])) & (~((D[3] & D[1]) & ~(D[4])) | D[8])) & (~((~(D[3]) & ~(D[1])) & D[4]) | D[6])) & (~((D[3] & ~(D[1])) & D[4]) | D[10])) & (~((~(D[3]) & D[1]) & D[4]) | D[11])) & (~((D[3] & D[1]) & D[4]) | D[9])

*)

FUNCTION_BLOCK F_CollectInput
  VAR_IN_OUT
      Data : ARRAY[1..15] OF BOOL;
  END_VAR
  VAR_INPUT
      TICK  : BOOL := 0;
      IN1   : BOOL := 0;
      IN2   : BOOL := 0;
      IN3   : BOOL := 0;
      IN4   : BOOL := 0;
      IN5   : BOOL := 0;
      RESET : BOOL := FALSE;
  END_VAR
  VAR_OUTPUT
      Finished : BOOL;
  END_VAR
  VAR
      j    : USINT := 1;
      tock : BOOL  := 0;
  END_VAR
  IF NOT RESET AND tock = NOT TICK THEN
      Data[j]   := IN1;
      Data[j+1] := IN2;
      Data[j+2] := IN3;
      Data[j+3] := IN4;
      Data[j+4] := IN5;
      j := j + 5;
      tock := TICK;
  ELSE
      j := 1;
      tock := 0;
  END_IF;
  Finished := (j > 15);
END_FUNCTION_BLOCK

PROGRAM Boiler
  VAR
    Data  : ARRAY[1..15] OF BOOL;
    Ready : BOOL;
    CollectInput : F_CollectInput;
  END_VAR
  VAR
    TICK     AT %IX1.0 : BOOL;
    IN1      AT %IX0.3 : BOOL;
    IN2      AT %IX0.4 : BOOL;
    IN3      AT %IX0.5 : BOOL;
    IN4      AT %IX0.6 : BOOL;
    IN5      AT %IX0.7 : BOOL;
    OutReady AT %QX0.0 : BOOL := FALSE;
    FeedNext AT %QX0.1 : BOOL := FALSE;
    Out      AT %QX0.2 : BOOL;
  END_VAR
  CollectInput(TICK:=TICK, IN1:=IN1, IN2:=IN2, IN3:=IN3, IN4:=IN4, IN5:=IN5);
  Ready := CollectInput.Finished;
  FeedNext := 1;
  IF Ready THEN
    Out := (((((((((NOT (((NOT D[3]) AND (NOT D[1])) AND (NOT D[4]))) OR D[5]) AND ((NOT ((D[3] AND (NOT D[1])) AND (NOT D[4]))) OR D[2])) AND ((NOT (((NOT D[3]) AND D[1]) AND (NOT D[4]))) OR D[7])) AND ((NOT ((D[3] AND D[1]) AND (NOT D[4]))) OR D[8])) AND ((NOT (((NOT D[3]) AND (NOT D[1])) AND D[4])) OR D[6])) AND ((NOT ((D[3] AND (NOT D[1])) AND D[4])) OR D[10])) AND ((NOT (((NOT D[3]) AND D[1]) AND D[4])) OR D[11])) AND ((NOT ((D[3] AND D[1]) AND D[4])) OR D[9]));
    OutReady := 1;
    CollectInput(RESET:=TRUE);
  END_IF;
END_PROGRAM

CONFIGURATION Config0
  RESOURCE Res0 ON PLC
    TASK task0(INTERVAL := T#20ms,PRIORITY := 0);
    PROGRAM instance0 WITH task0 : Boiler;
  END_RESOURCE
END_CONFIGURATION

(* ---- 3-MUX_plebe-tasks-woozy.st ---- *)
(*
This code implements a shuffled multiplexer with 3 control bits.
The control bits are: Data[2], Data[1], Data[3]
The input bits are: Data[8], Data[6], Data[7], Data[5], Data[9], Data[4], Data[10], Data[11]

The symbolic expression is:
(((((((~((~(D[2]) & ~(D[1])) & ~(D[3])) | D[8]) & (~((D[2] & ~(D[1])) & ~(D[3])) | D[6])) & (~((~(D[2]) & D[1]) & ~(D[3])) | D[7])) & (~((D[2] & D[1]) & ~(D[3])) | D[5])) & (~((~(D[2]) & ~(D[1])) & D[3]) | D[9])) & (~((D[2] & ~(D[1])) & D[3]) | D[4])) & (~((~(D[2]) & D[1]) & D[3]) | D[10])) & (~((D[2] & D[1]) & D[3]) | D[11])

*)

FUNCTION_BLOCK F_CollectInput
  VAR_IN_OUT
      Data : ARRAY[1..15] OF BOOL;
  END_VAR
  VAR_INPUT
      TICK  : BOOL := 0;
      IN1   : BOOL := 0;
      IN2   : BOOL := 0;
      IN3   : BOOL := 0;
      IN4   : BOOL := 0;
      IN5   : BOOL := 0;
      RESET : BOOL := FALSE;
  END_VAR
  VAR_OUTPUT
      Finished : BOOL;
  END_VAR
  VAR
      j    : USINT := 1;
      tock : BOOL  := 0;
  END_VAR
  IF NOT RESET AND tock = NOT TICK THEN
      Data[j]   := IN1;
      Data[j+1] := IN2;
      Data[j+2] := IN3;
      Data[j+3] := IN4;
      Data[j+4] := IN5;
      j := j + 5;
      tock := TICK;
  ELSE
      j := 1;
      tock := 0;
  END_IF;
  Finished := (j > 15);
END_FUNCTION_BLOCK

PROGRAM Boiler
  VAR
    Data  : ARRAY[1..15] OF BOOL;
    Ready : BOOL;
    CollectInput : F_CollectInput;
  END_VAR
  VAR
    TICK     AT %IX1.0 : BOOL;
    IN1      AT %IX0.3 : BOOL;
    IN2      AT %IX0.4 : BOOL;
    IN3      AT %IX0.5 : BOOL;
    IN4      AT %IX0.6 : BOOL;
    IN5      AT %IX0.7 : BOOL;
    OutReady AT %QX0.0 : BOOL := FALSE;
    FeedNext AT %QX0.1 : BOOL := FALSE;
    Out      AT %QX0.2 : BOOL;
  END_VAR
  CollectInput(TICK:=TICK, IN1:=IN1, IN2:=IN2, IN3:=IN3, IN4:=IN4, IN5:=IN5);
  Ready := CollectInput.Finished;
  FeedNext := 1;
  IF Ready THEN
    Out := (((((((((NOT (((NOT D[2]) AND (NOT D[1])) AND (NOT D[3]))) OR D[8]) AND ((NOT ((D[2] AND (NOT D[1])) AND (NOT D[3]))) OR D[6])) AND ((NOT (((NOT D[2]) AND D[1]) AND (NOT D[3]))) OR D[7])) AND ((NOT ((D[2] AND D[1]) AND (NOT D[3]))) OR D[5])) AND ((NOT (((NOT D[2]) AND (NOT D[1])) AND D[3])) OR D[9])) AND ((NOT ((D[2] AND (NOT D[1])) AND D[3])) OR D[4])) AND ((NOT (((NOT D[2]) AND D[1]) AND D[3])) OR D[10])) AND ((NOT ((D[2] AND D[1]) AND D[3])) OR D[11]));
    OutReady := 1;
    CollectInput(RESET:=TRUE);
  END_IF;
END_PROGRAM

CONFIGURATION Config0
  RESOURCE Res0 ON PLC
    TASK task0(INTERVAL := T#20ms,PRIORITY := 0);
    PROGRAM instance0 WITH task0 : Boiler;
  END_RESOURCE
END_CONFIGURATION

(* ---- 3-MUX_poser-hayer-swain.st ---- *)
(*
This code implements a shuffled multiplexer with 3 control bits.
The control bits are: Data[9], Data[2], Data[3]
The input bits are: Data[4], Data[1], Data[5], Data[10], Data[11], Data[8], Data[7], Data[6]

The symbolic expression is:
(((((((~((~(D[9]) & ~(D[2])) & ~(D[3])) | D[4]) & (~((D[9] & ~(D[2])) & ~(D[3])) | D[1])) & (~((~(D[9]) & D[2]) & ~(D[3])) | D[5])) & (~((D[9] & D[2]) & ~(D[3])) | D[10])) & (~((~(D[9]) & ~(D[2])) & D[3]) | D[11])) & (~((D[9] & ~(D[2])) & D[3]) | D[8])) & (~((~(D[9]) & D[2]) & D[3]) | D[7])) & (~((D[9] & D[2]) & D[3]) | D[6])

*)

FUNCTION_BLOCK F_CollectInput
  VAR_IN_OUT
      Data : ARRAY[1..15] OF BOOL;
  END_VAR
  VAR_INPUT
      TICK  : BOOL := 0;
      IN1   : BOOL := 0;
      IN2   : BOOL := 0;
      IN3   : BOOL := 0;
      IN4   : BOOL := 0;
      IN5   : BOOL := 0;
      RESET : BOOL := FALSE;
  END_VAR
  VAR_OUTPUT
      Finished : BOOL;
  END_VAR
  VAR
      j    : USINT := 1;
      tock : BOOL  := 0;
  END_VAR
  IF NOT RESET AND tock = NOT TICK THEN
      Data[j]   := IN1;
      Data[j+1] := IN2;
      Data[j+2] := IN3;
      Data[j+3] := IN4;
      Data[j+4] := IN5;
      j := j + 5;
      tock := TICK;
  ELSE
      j := 1;
      tock := 0;
  END_IF;
  Finished := (j > 15);
END_FUNCTION_BLOCK

PROGRAM Boiler
  VAR
    Data  : ARRAY[1..15] OF BOOL;
    Ready : BOOL;
    CollectInput : F_CollectInput;
  END_VAR
  VAR
    TICK     AT %IX1.0 : BOOL;
    IN1      AT %IX0.3 : BOOL;
    IN2      AT %IX0.4 : BOOL;
    IN3      AT %IX0.5 : BOOL;
    IN4      AT %IX0.6 : BOOL;
    IN5      AT %IX0.7 : BOOL;
    OutReady AT %QX0.0 : BOOL := FALSE;
    FeedNext AT %QX0.1 : BOOL := FALSE;
    Out      AT %QX0.2 : BOOL;
  END_VAR
  CollectInput(TICK:=TICK, IN1:=IN1, IN2:=IN2, IN3:=IN3, IN4:=IN4, IN5:=IN5);
  Ready := CollectInput.Finished;
  FeedNext := 1;
  IF Ready THEN
    Out := (((((((((NOT (((NOT D[9]) AND (NOT D[2])) AND (NOT D[3]))) OR D[4]) AND ((NOT ((D[9] AND (NOT D[2])) AND (NOT D[3]))) OR D[1])) AND ((NOT (((NOT D[9]) AND D[2]) AND (NOT D[3]))) OR D[5])) AND ((NOT ((D[9] AND D[2]) AND (NOT D[3]))) OR D[10])) AND ((NOT (((NOT D[9]) AND (NOT D[2])) AND D[3])) OR D[11])) AND ((NOT ((D[9] AND (NOT D[2])) AND D[3])) OR D[8])) AND ((NOT (((NOT D[9]) AND D[2]) AND D[3])) OR D[7])) AND ((NOT ((D[9] AND D[2]) AND D[3])) OR D[6]));
    OutReady := 1;
    CollectInput(RESET:=TRUE);
  END_IF;
END_PROGRAM

CONFIGURATION Config0
  RESOURCE Res0 ON PLC
    TASK task0(INTERVAL := T#20ms,PRIORITY := 0);
    PROGRAM instance0 WITH task0 : Boiler;
  END_RESOURCE
END_CONFIGURATION

(* ---- 3-MUX_pseud-hurts-novas.st ---- *)
(*
This code implements a shuffled multiplexer with 3 control bits.
The control bits are: Data[3], Data[1], Data[2]
The input bits are: Data[4], Data[5], Data[10], Data[9], Data[7], Data[8], Data[11], Data[6]

The symbolic expression is:
(((((((~((~(D[3]) & ~(D[1])) & ~(D[2])) | D[4]) & (~((D[3] & ~(D[1])) & ~(D[2])) | D[5])) & (~((~(D[3]) & D[1]) & ~(D[2])) | D[10])) & (~((D[3] & D[1]) & ~(D[2])) | D[9])) & (~((~(D[3]) & ~(D[1])) & D[2]) | D[7])) & (~((D[3] & ~(D[1])) & D[2]) | D[8])) & (~((~(D[3]) & D[1]) & D[2]) | D[11])) & (~((D[3] & D[1]) & D[2]) | D[6])

*)

FUNCTION_BLOCK F_CollectInput
  VAR_IN_OUT
      Data : ARRAY[1..15] OF BOOL;
  END_VAR
  VAR_INPUT
      TICK  : BOOL := 0;
      IN1   : BOOL := 0;
      IN2   : BOOL := 0;
      IN3   : BOOL := 0;
      IN4   : BOOL := 0;
      IN5   : BOOL := 0;
      RESET : BOOL := FALSE;
  END_VAR
  VAR_OUTPUT
      Finished : BOOL;
  END_VAR
  VAR
      j    : USINT := 1;
      tock : BOOL  := 0;
  END_VAR
  IF NOT RESET AND tock = NOT TICK THEN
      Data[j]   := IN1;
      Data[j+1] := IN2;
      Data[j+2] := IN3;
      Data[j+3] := IN4;
      Data[j+4] := IN5;
      j := j + 5;
      tock := TICK;
  ELSE
      j := 1;
      tock := 0;
  END_IF;
  Finished := (j > 15);
END_FUNCTION_BLOCK

PROGRAM Boiler
  VAR
    Data  : ARRAY[1..15] OF BOOL;
    Ready : BOOL;
    CollectInput : F_CollectInput;
  END_VAR
  VAR
    TICK     AT %IX1.0 : BOOL;
    IN1      AT %IX0.3 : BOOL;
    IN2      AT %IX0.4 : BOOL;
    IN3      AT %IX0.5 : BOOL;
    IN4      AT %IX0.6 : BOOL;
    IN5      AT %IX0.7 : BOOL;
    OutReady AT %QX0.0 : BOOL := FALSE;
    FeedNext AT %QX0.1 : BOOL := FALSE;
    Out      AT %QX0.2 : BOOL;
  END_VAR
  CollectInput(TICK:=TICK, IN1:=IN1, IN2:=IN2, IN3:=IN3, IN4:=IN4, IN5:=IN5);
  Ready := CollectInput.Finished;
  FeedNext := 1;
  IF Ready THEN
    Out := (((((((((NOT (((NOT D[3]) AND (NOT D[1])) AND (NOT D[2]))) OR D[4]) AND ((NOT ((D[3] AND (NOT D[1])) AND (NOT D[2]))) OR D[5])) AND ((NOT (((NOT D[3]) AND D[1]) AND (NOT D[2]))) OR D[10])) AND ((NOT ((D[3] AND D[1]) AND (NOT D[2]))) OR D[9])) AND ((NOT (((NOT D[3]) AND (NOT D[1])) AND D[2])) OR D[7])) AND ((NOT ((D[3] AND (NOT D[1])) AND D[2])) OR D[8])) AND ((NOT (((NOT D[3]) AND D[1]) AND D[2])) OR D[11])) AND ((NOT ((D[3] AND D[1]) AND D[2])) OR D[6]));
    OutReady := 1;
    CollectInput(RESET:=TRUE);
  END_IF;
END_PROGRAM

CONFIGURATION Config0
  RESOURCE Res0 ON PLC
    TASK task0(INTERVAL := T#20ms,PRIORITY := 0);
    PROGRAM instance0 WITH task0 : Boiler;
  END_RESOURCE
END_CONFIGURATION

(* ---- 3-MUX_quire-amigo-polis.st ---- *)
(*
This code implements a shuffled multiplexer with 3 control bits.
The control bits are: Data[1], Data[2], Data[4]
The input bits are: Data[5], Data[9], Data[6], Data[11], Data[7], Data[3], Data[10], Data[8]

The symbolic expression is:
(((((((~((~(D[1]) & ~(D[2])) & ~(D[4])) | D[5]) & (~((D[1] & ~(D[2])) & ~(D[4])) | D[9])) & (~((~(D[1]) & D[2]) & ~(D[4])) | D[6])) & (~((D[1] & D[2]) & ~(D[4])) | D[11])) & (~((~(D[1]) & ~(D[2])) & D[4]) | D[7])) & (~((D[1] & ~(D[2])) & D[4]) | D[3])) & (~((~(D[1]) & D[2]) & D[4]) | D[10])) & (~((D[1] & D[2]) & D[4]) | D[8])

*)

FUNCTION_BLOCK F_CollectInput
  VAR_IN_OUT
      Data : ARRAY[1..15] OF BOOL;
  END_VAR
  VAR_INPUT
      TICK  : BOOL := 0;
      IN1   : BOOL := 0;
      IN2   : BOOL := 0;
      IN3   : BOOL := 0;
      IN4   : BOOL := 0;
      IN5   : BOOL := 0;
      RESET : BOOL := FALSE;
  END_VAR
  VAR_OUTPUT
      Finished : BOOL;
  END_VAR
  VAR
      j    : USINT := 1;
      tock : BOOL  := 0;
  END_VAR
  IF NOT RESET AND tock = NOT TICK THEN
      Data[j]   := IN1;
      Data[j+1] := IN2;
      Data[j+2] := IN3;
      Data[j+3] := IN4;
      Data[j+4] := IN5;
      j := j + 5;
      tock := TICK;
  ELSE
      j := 1;
      tock := 0;
  END_IF;
  Finished := (j > 15);
END_FUNCTION_BLOCK

PROGRAM Boiler
  VAR
    Data  : ARRAY[1..15] OF BOOL;
    Ready : BOOL;
    CollectInput : F_CollectInput;
  END_VAR
  VAR
    TICK     AT %IX1.0 : BOOL;
    IN1      AT %IX0.3 : BOOL;
    IN2      AT %IX0.4 : BOOL;
    IN3      AT %IX0.5 : BOOL;
    IN4      AT %IX0.6 : BOOL;
    IN5      AT %IX0.7 : BOOL;
    OutReady AT %QX0.0 : BOOL := FALSE;
    FeedNext AT %QX0.1 : BOOL := FALSE;
    Out      AT %QX0.2 : BOOL;
  END_VAR
  CollectInput(TICK:=TICK, IN1:=IN1, IN2:=IN2, IN3:=IN3, IN4:=IN4, IN5:=IN5);
  Ready := CollectInput.Finished;
  FeedNext := 1;
  IF Ready THEN
    Out := (((((((((NOT (((NOT D[1]) AND (NOT D[2])) AND (NOT D[4]))) OR D[5]) AND ((NOT ((D[1] AND (NOT D[2])) AND (NOT D[4]))) OR D[9])) AND ((NOT (((NOT D[1]) AND D[2]) AND (NOT D[4]))) OR D[6])) AND ((NOT ((D[1] AND D[2]) AND (NOT D[4]))) OR D[11])) AND ((NOT (((NOT D[1]) AND (NOT D[2])) AND D[4])) OR D[7])) AND ((NOT ((D[1] AND (NOT D[2])) AND D[4])) OR D[3])) AND ((NOT (((NOT D[1]) AND D[2]) AND D[4])) OR D[10])) AND ((NOT ((D[1] AND D[2]) AND D[4])) OR D[8]));
    OutReady := 1;
    CollectInput(RESET:=TRUE);
  END_IF;
END_PROGRAM

CONFIGURATION Config0
  RESOURCE Res0 ON PLC
    TASK task0(INTERVAL := T#20ms,PRIORITY := 0);
    PROGRAM instance0 WITH task0 : Boiler;
  END_RESOURCE
END_CONFIGURATION

(* ---- 3-MUX_reign-bends-kebob.st ---- *)
(*
This code implements a shuffled multiplexer with 3 control bits.
The control bits are: Data[6], Data[3], Data[4]
The input bits are: Data[2], Data[1], Data[5], Data[7], Data[9], Data[8], Data[10], Data[11]

The symbolic expression is:
(((((((~((~(D[6]) & ~(D[3])) & ~(D[4])) | D[2]) & (~((D[6] & ~(D[3])) & ~(D[4])) | D[1])) & (~((~(D[6]) & D[3]) & ~(D[4])) | D[5])) & (~((D[6] & D[3]) & ~(D[4])) | D[7])) & (~((~(D[6]) & ~(D[3])) & D[4]) | D[9])) & (~((D[6] & ~(D[3])) & D[4]) | D[8])) & (~((~(D[6]) & D[3]) & D[4]) | D[10])) & (~((D[6] & D[3]) & D[4]) | D[11])

*)

FUNCTION_BLOCK F_CollectInput
  VAR_IN_OUT
      Data : ARRAY[1..15] OF BOOL;
  END_VAR
  VAR_INPUT
      TICK  : BOOL := 0;
      IN1   : BOOL := 0;
      IN2   : BOOL := 0;
      IN3   : BOOL := 0;
      IN4   : BOOL := 0;
      IN5   : BOOL := 0;
      RESET : BOOL := FALSE;
  END_VAR
  VAR_OUTPUT
      Finished : BOOL;
  END_VAR
  VAR
      j    : USINT := 1;
      tock : BOOL  := 0;
  END_VAR
  IF NOT RESET AND tock = NOT TICK THEN
      Data[j]   := IN1;
      Data[j+1] := IN2;
      Data[j+2] := IN3;
      Data[j+3] := IN4;
      Data[j+4] := IN5;
      j := j + 5;
      tock := TICK;
  ELSE
      j := 1;
      tock := 0;
  END_IF;
  Finished := (j > 15);
END_FUNCTION_BLOCK

PROGRAM Boiler
  VAR
    Data  : ARRAY[1..15] OF BOOL;
    Ready : BOOL;
    CollectInput : F_CollectInput;
  END_VAR
  VAR
    TICK     AT %IX1.0 : BOOL;
    IN1      AT %IX0.3 : BOOL;
    IN2      AT %IX0.4 : BOOL;
    IN3      AT %IX0.5 : BOOL;
    IN4      AT %IX0.6 : BOOL;
    IN5      AT %IX0.7 : BOOL;
    OutReady AT %QX0.0 : BOOL := FALSE;
    FeedNext AT %QX0.1 : BOOL := FALSE;
    Out      AT %QX0.2 : BOOL;
  END_VAR
  CollectInput(TICK:=TICK, IN1:=IN1, IN2:=IN2, IN3:=IN3, IN4:=IN4, IN5:=IN5);
  Ready := CollectInput.Finished;
  FeedNext := 1;
  IF Ready THEN
    Out := (((((((((NOT (((NOT D[6]) AND (NOT D[3])) AND (NOT D[4]))) OR D[2]) AND ((NOT ((D[6] AND (NOT D[3])) AND (NOT D[4]))) OR D[1])) AND ((NOT (((NOT D[6]) AND D[3]) AND (NOT D[4]))) OR D[5])) AND ((NOT ((D[6] AND D[3]) AND (NOT D[4]))) OR D[7])) AND ((NOT (((NOT D[6]) AND (NOT D[3])) AND D[4])) OR D[9])) AND ((NOT ((D[6] AND (NOT D[3])) AND D[4])) OR D[8])) AND ((NOT (((NOT D[6]) AND D[3]) AND D[4])) OR D[10])) AND ((NOT ((D[6] AND D[3]) AND D[4])) OR D[11]));
    OutReady := 1;
    CollectInput(RESET:=TRUE);
  END_IF;
END_PROGRAM

CONFIGURATION Config0
  RESOURCE Res0 ON PLC
    TASK task0(INTERVAL := T#20ms,PRIORITY := 0);
    PROGRAM instance0 WITH task0 : Boiler;
  END_RESOURCE
END_CONFIGURATION
